(* IEC 61131-3 sources: Aqueous_Solutions/docs-authority/plc, 18 files *)

(* ---- PLC-CRYO.st ---- *)
(* AQS-CTL-004 X-CTL-04: control program source, generated by flow_graph/control/plc_programs.py *)
(* Basis: AQS-CTL-001 INSTRUMENT_INDEX.csv, AQS-CTL-002 control architecture, graph set-points. *)
(* PLC-CRYO: CPU redundant pair; IO counts AI 36 AO 1 DI 19 DO 6 (modules per AQS-CTL-002, 16-channel, 20 % spare) *)
PROGRAM PLC_CRYO_CTRL
VAR
  (* 100 ms cyclic task per AQS-CTL-002 *)
  CRYO_AHU_COND_CONDENSABLEFT-01_PV : REAL ;  (* S70 normal 0.00 L/h )
  CRYO_AHU_COND_CONDENSABLEPT-01_PV : REAL ;  (* no design pressure on the graph )
  CRYO_AHU_COND_CONDENSABLETE-01_PV : REAL ;  (* band by service )
  CRYO_AHUFT-01_PV : REAL ;  (* S56 normal 0.00 L/h )
  CRYO_AHUFT-02_PV : REAL ;  (* S68 normal 4.27 L/h )
  CRYO_AHUFT-03_PV : REAL ;  (* S86 normal 0.00 L/h )
  CRYO_AHUFT-04_PV : REAL ;  (* IA-HVAC-COND normal 2.81 L/h )
  CRYO_AHUPT-01_PV : REAL ;  (* no design pressure on the graph )
  CRYO_AHUTE-01_PV : REAL ;  (* band by service )
  CRYO_ASUPT-01_PV : REAL ;  (* design 18.0 kPa g )
  CRYO_ASUTE-01_PV : REAL ;  (* band by service )
  CRYO_CO2PT-01_PV : REAL ;  (* design 2200.0 kPa g )
  CRYO_CO2TE-01_PV : REAL ;  (* design T 25 C )
  CRYO_DED_COOLPT-01_PV : REAL ;  (* no design pressure on the graph )
  CRYO_DED_COOLTE-01_PV : REAL ;  (* band by service )
  CRYO_H2PT-01_PV : REAL ;  (* design 22000.0 kPa g )
  CRYO_H2TE-01_PV : REAL ;  (* design T 25 C )
  CRYO_N2PT-01_PV : REAL ;  (* no design pressure on the graph )
  CRYO_N2TE-01_PV : REAL ;  (* band by service )
  CRYO_O2PT-01_PV : REAL ;  (* design 22000.0 kPa g )
  CRYO_O2TE-01_PV : REAL ;  (* design T 25 C )
  CRYO_HX_Q4PT-01_PV : REAL ;  (* no design pressure on the graph )
  CRYO_HX_Q4TE-01_PV : REAL ;  (* band by service )
  H2O_ELYZFT-01_PV : REAL ;  (* IA-ELY-H2 normal 0.43 L/h )
  H2O_ELYZFT-02_PV : REAL ;  (* IA-ELY-O2 normal 3.42 L/h )
  H2O_ELYZLT-01_PV : REAL ;  (* A-M-182 liquid height )
  H2O_ELYZPT-01_PV : REAL ;  (* design 990.0 kPa g )
  H2O_ELYZTE-01_PV : REAL ;  (* band by service )
  PROD_MEOHLT-01_PV : REAL ;  (* A-M-182 liquid height )
  PROD_MEOHPT-01_PV : REAL ;  (* no design pressure on the graph )
  PROD_MEOHTE-01_PV : REAL ;  (* band by service )
  PROD_O2PT-01_PV : REAL ;  (* no design pressure on the graph )
  PROD_O2TE-01_PV : REAL ;  (* band by service )
  AIR_RECEIVERPT-01_PV : REAL ;  (* no design pressure on the graph )
  AIR_RECEIVERTE-01_PV : REAL ;  (* band by service )
  PROD_MEOHFT-01_PV : REAL ;  (* methanol product: IA-MEOH-PROD 28.15 kg/d (1.50 L/h at 792 kg/m3) )
END_VAR

  (* FLOW control loop - set-point from the graph basis *)
  CRYO_AHU_COND_CONDENSABLEFT-01_SP := 0.0 ;  (* graph basis: S70 normal 0.00 L/h )
  FB_PI_CRYO_AHU_COND_CONDENSABLEFT-01( PV := CRYO_AHU_COND_CONDENSABLEFT-01_PV, SP := CRYO_AHU_COND_CONDENSABLEFT-01_SP );  (* PI per AQS-CTL-002; GAIN/KI entered at commissioning from the step test (AQS-COM-001 sec. 3), anti-windup clamp per this FB *)
  CRYO_AHU_COND_CONDENSABLEFT-01_ALARM_HI := 0.0 ;  (* expected-zero state: any positive PV alarms )

  (* PRESSURE monitoring block - indication, no set-point invented )
  FB_AI_CRYO_AHU_COND_CONDENSABLEPT-01( PV := CRYO_AHU_COND_CONDENSABLEPT-01_PV );
  CRYO_AHU_COND_CONDENSABLEPT-01_ALARM_HI := 9.0 ;  (* 90 % of span, registered LSH convention )

  (* TEMPERATURE monitoring block - indication, no set-point invented )
  FB_AI_CRYO_AHU_COND_CONDENSABLETE-01( PV := CRYO_AHU_COND_CONDENSABLETE-01_PV );
  CRYO_AHU_COND_CONDENSABLETE-01_ALARM_HI := 45.0 ;  (* 90 % of span, registered LSH convention )

  (* FLOW control loop - set-point from the graph basis *)
  CRYO_AHUFT-01_SP := 0.0 ;  (* graph basis: S56 normal 0.00 L/h )
  FB_PI_CRYO_AHUFT-01( PV := CRYO_AHUFT-01_PV, SP := CRYO_AHUFT-01_SP );  (* PI per AQS-CTL-002; GAIN/KI entered at commissioning from the step test (AQS-COM-001 sec. 3), anti-windup clamp per this FB *)
  CRYO_AHUFT-01_ALARM_HI := 0.0 ;  (* expected-zero state: any positive PV alarms )

  (* FLOW control loop - set-point from the graph basis *)
  CRYO_AHUFT-02_SP := 4.27 ;  (* graph basis: S68 normal 4.27 L/h )
  FB_PI_CRYO_AHUFT-02( PV := CRYO_AHUFT-02_PV, SP := CRYO_AHUFT-02_SP );  (* PI per AQS-CTL-002; GAIN/KI entered at commissioning from the step test (AQS-COM-001 sec. 3), anti-windup clamp per this FB *)
  CRYO_AHUFT-02_ALARM_HI := 4.697 ;  (* SP x 1.1 margin, A-M-188 margin class *)
  CRYO_AHUFT-02_ALARM_LO := 3.8429999999999995 ;

  (* FLOW control loop - set-point from the graph basis *)
  CRYO_AHUFT-03_SP := 0.0 ;  (* graph basis: S86 normal 0.00 L/h )
  FB_PI_CRYO_AHUFT-03( PV := CRYO_AHUFT-03_PV, SP := CRYO_AHUFT-03_SP );  (* PI per AQS-CTL-002; GAIN/KI entered at commissioning from the step test (AQS-COM-001 sec. 3), anti-windup clamp per this FB *)
  CRYO_AHUFT-03_ALARM_HI := 0.0 ;  (* expected-zero state: any positive PV alarms )

  (* FLOW control loop - set-point from the graph basis *)
  CRYO_AHUFT-04_SP := 2.81 ;  (* graph basis: IA-HVAC-COND normal 2.81 L/h )
  FB_PI_CRYO_AHUFT-04( PV := CRYO_AHUFT-04_PV, SP := CRYO_AHUFT-04_SP );  (* PI per AQS-CTL-002; GAIN/KI entered at commissioning from the step test (AQS-COM-001 sec. 3), anti-windup clamp per this FB *)
  CRYO_AHUFT-04_ALARM_HI := 3.091 ;  (* SP x 1.1 margin, A-M-188 margin class *)
  CRYO_AHUFT-04_ALARM_LO := 2.529 ;

  (* PRESSURE monitoring block - indication, no set-point invented )
  FB_AI_CRYO_AHUPT-01( PV := CRYO_AHUPT-01_PV );
  CRYO_AHUPT-01_ALARM_HI := 9.0 ;  (* 90 % of span, registered LSH convention )

  (* TEMPERATURE monitoring block - indication, no set-point invented )
  FB_AI_CRYO_AHUTE-01( PV := CRYO_AHUTE-01_PV );
  CRYO_AHUTE-01_ALARM_HI := 45.0 ;  (* 90 % of span, registered LSH convention )

  (* PRESSURE control loop - set-point from the graph basis *)
  CRYO_ASUPT-01_SP := 18.0 ;  (* graph basis: design 18.0 kPa g )
  FB_PI_CRYO_ASUPT-01( PV := CRYO_ASUPT-01_PV, SP := CRYO_ASUPT-01_SP );  (* PI per AQS-CTL-002; GAIN/KI entered at commissioning from the step test (AQS-COM-001 sec. 3), anti-windup clamp per this FB *)
  CRYO_ASUPT-01_ALARM_HI := 19.8 ;  (* SP x 1.1 margin, A-M-188 margin class *)
  CRYO_ASUPT-01_ALARM_LO := 16.2 ;

  (* TEMPERATURE monitoring block - indication, no set-point invented )
  FB_AI_CRYO_ASUTE-01( PV := CRYO_ASUTE-01_PV );
  CRYO_ASUTE-01_ALARM_HI := 45.0 ;  (* 90 % of span, registered LSH convention )

  (* PRESSURE control loop - set-point from the graph basis *)
  CRYO_CO2PT-01_SP := 2200.0 ;  (* graph basis: design 2200.0 kPa g )
  FB_PI_CRYO_CO2PT-01( PV := CRYO_CO2PT-01_PV, SP := CRYO_CO2PT-01_SP );  (* PI per AQS-CTL-002; GAIN/KI entered at commissioning from the step test (AQS-COM-001 sec. 3), anti-windup clamp per this FB *)
  CRYO_CO2PT-01_ALARM_HI := 2420.0 ;  (* SP x 1.1 margin, A-M-188 margin class *)
  CRYO_CO2PT-01_ALARM_LO := 1980.0 ;

  (* TEMPERATURE control loop - set-point from the graph basis *)
  CRYO_CO2TE-01_SP := 25.0 ;  (* graph basis: design T 25 C )
  FB_PI_CRYO_CO2TE-01( PV := CRYO_CO2TE-01_PV, SP := CRYO_CO2TE-01_SP );  (* PI per AQS-CTL-002; GAIN/KI entered at commissioning from the step test (AQS-COM-001 sec. 3), anti-windup clamp per this FB *)
  CRYO_CO2TE-01_ALARM_HI := 27.500000000000004 ;  (* SP x 1.1 margin, A-M-188 margin class *)
  CRYO_CO2TE-01_ALARM_LO := 22.5 ;

  (* PRESSURE monitoring block - indication, no set-point invented )
  FB_AI_CRYO_DED_COOLPT-01( PV := CRYO_DED_COOLPT-01_PV );
  CRYO_DED_COOLPT-01_ALARM_HI := 9.0 ;  (* 90 % of span, registered LSH convention )

  (* TEMPERATURE monitoring block - indication, no set-point invented )
  FB_AI_CRYO_DED_COOLTE-01( PV := CRYO_DED_COOLTE-01_PV );
  CRYO_DED_COOLTE-01_ALARM_HI := 45.0 ;  (* 90 % of span, registered LSH convention )

  (* PRESSURE control loop - set-point from the graph basis *)
  CRYO_H2PT-01_SP := 22000.0 ;  (* graph basis: design 22000.0 kPa g )
  FB_PI_CRYO_H2PT-01( PV := CRYO_H2PT-01_PV, SP := CRYO_H2PT-01_SP );  (* PI per AQS-CTL-002; GAIN/KI entered at commissioning from the step test (AQS-COM-001 sec. 3), anti-windup clamp per this FB *)
  CRYO_H2PT-01_ALARM_HI := 24200.000000000004 ;  (* SP x 1.1 margin, A-M-188 margin class *)
  CRYO_H2PT-01_ALARM_LO := 19800.0 ;

  (* TEMPERATURE control loop - set-point from the graph basis *)
  CRYO_H2TE-01_SP := 25.0 ;  (* graph basis: design T 25 C )
  FB_PI_CRYO_H2TE-01( PV := CRYO_H2TE-01_PV, SP := CRYO_H2TE-01_SP );  (* PI per AQS-CTL-002; GAIN/KI entered at commissioning from the step test (AQS-COM-001 sec. 3), anti-windup clamp per this FB *)
  CRYO_H2TE-01_ALARM_HI := 27.500000000000004 ;  (* SP x 1.1 margin, A-M-188 margin class *)
  CRYO_H2TE-01_ALARM_LO := 22.5 ;

  (* PRESSURE monitoring block - indication, no set-point invented )
  FB_AI_CRYO_N2PT-01( PV := CRYO_N2PT-01_PV );
  CRYO_N2PT-01_ALARM_HI := 9.0 ;  (* 90 % of span, registered LSH convention )

  (* TEMPERATURE monitoring block - indication, no set-point invented )
  FB_AI_CRYO_N2TE-01( PV := CRYO_N2TE-01_PV );
  CRYO_N2TE-01_ALARM_HI := 45.0 ;  (* 90 % of span, registered LSH convention )

  (* PRESSURE control loop - set-point from the graph basis *)
  CRYO_O2PT-01_SP := 22000.0 ;  (* graph basis: design 22000.0 kPa g )
  FB_PI_CRYO_O2PT-01( PV := CRYO_O2PT-01_PV, SP := CRYO_O2PT-01_SP );  (* PI per AQS-CTL-002; GAIN/KI entered at commissioning from the step test (AQS-COM-001 sec. 3), anti-windup clamp per this FB *)
  CRYO_O2PT-01_ALARM_HI := 24200.000000000004 ;  (* SP x 1.1 margin, A-M-188 margin class *)
  CRYO_O2PT-01_ALARM_LO := 19800.0 ;

  (* TEMPERATURE control loop - set-point from the graph basis *)
  CRYO_O2TE-01_SP := 25.0 ;  (* graph basis: design T 25 C )
  FB_PI_CRYO_O2TE-01( PV := CRYO_O2TE-01_PV, SP := CRYO_O2TE-01_SP );  (* PI per AQS-CTL-002; GAIN/KI entered at commissioning from the step test (AQS-COM-001 sec. 3), anti-windup clamp per this FB *)
  CRYO_O2TE-01_ALARM_HI := 27.500000000000004 ;  (* SP x 1.1 margin, A-M-188 margin class *)
  CRYO_O2TE-01_ALARM_LO := 22.5 ;

  (* PRESSURE monitoring block - indication, no set-point invented )
  FB_AI_CRYO_HX_Q4PT-01( PV := CRYO_HX_Q4PT-01_PV );
  CRYO_HX_Q4PT-01_ALARM_HI := 9.0 ;  (* 90 % of span, registered LSH convention )

  (* TEMPERATURE monitoring block - indication, no set-point invented )
  FB_AI_CRYO_HX_Q4TE-01( PV := CRYO_HX_Q4TE-01_PV );
  CRYO_HX_Q4TE-01_ALARM_HI := 45.0 ;  (* 90 % of span, registered LSH convention )

  (* FLOW control loop - set-point from the graph basis *)
  H2O_ELYZFT-01_SP := 0.43 ;  (* graph basis: IA-ELY-H2 normal 0.43 L/h )
  FB_PI_H2O_ELYZFT-01( PV := H2O_ELYZFT-01_PV, SP := H2O_ELYZFT-01_SP );  (* PI per AQS-CTL-002; GAIN/KI entered at commissioning from the step test (AQS-COM-001 sec. 3), anti-windup clamp per this FB *)
  H2O_ELYZFT-01_ALARM_HI := 0.47300000000000003 ;  (* SP x 1.1 margin, A-M-188 margin class *)
  H2O_ELYZFT-01_ALARM_LO := 0.387 ;

  (* FLOW control loop - set-point from the graph basis *)
  H2O_ELYZFT-02_SP := 3.42 ;  (* graph basis: IA-ELY-O2 normal 3.42 L/h )
  FB_PI_H2O_ELYZFT-02( PV := H2O_ELYZFT-02_PV, SP := H2O_ELYZFT-02_SP );  (* PI per AQS-CTL-002; GAIN/KI entered at commissioning from the step test (AQS-COM-001 sec. 3), anti-windup clamp per this FB *)
  H2O_ELYZFT-02_ALARM_HI := 3.762 ;  (* SP x 1.1 margin, A-M-188 margin class *)
  H2O_ELYZFT-02_ALARM_LO := 3.078 ;

  (* LEVEL monitoring block - indication, no set-point invented )
  FB_AI_H2O_ELYZLT-01( PV := H2O_ELYZLT-01_PV );
  H2O_ELYZLT-01_ALARM_HI := 90.0 ;  (* 90 % of span, registered LSH convention )

  (* PRESSURE control loop - set-point from the graph basis *)
  H2O_ELYZPT-01_SP := 990.0 ;  (* graph basis: design 990.0 kPa g )
  FB_PI_H2O_ELYZPT-01( PV := H2O_ELYZPT-01_PV, SP := H2O_ELYZPT-01_SP );  (* PI per AQS-CTL-002; GAIN/KI entered at commissioning from the step test (AQS-COM-001 sec. 3), anti-windup clamp per this FB *)
  H2O_ELYZPT-01_ALARM_HI := 1089.0 ;  (* SP x 1.1 margin, A-M-188 margin class *)
  H2O_ELYZPT-01_ALARM_LO := 891.0 ;

  (* TEMPERATURE monitoring block - indication, no set-point invented )
  FB_AI_H2O_ELYZTE-01( PV := H2O_ELYZTE-01_PV );
  H2O_ELYZTE-01_ALARM_HI := 135.0 ;  (* 90 % of span, registered LSH convention )

  (* LEVEL monitoring block - indication, no set-point invented )
  FB_AI_PROD_MEOHLT-01( PV := PROD_MEOHLT-01_PV );
  PROD_MEOHLT-01_ALARM_HI := 90.0 ;  (* 90 % of span, registered LSH convention )

  (* PRESSURE monitoring block - indication, no set-point invented )
  FB_AI_PROD_MEOHPT-01( PV := PROD_MEOHPT-01_PV );
  PROD_MEOHPT-01_ALARM_HI := 9.0 ;  (* 90 % of span, registered LSH convention )

  (* TEMPERATURE monitoring block - indication, no set-point invented )
  FB_AI_PROD_MEOHTE-01( PV := PROD_MEOHTE-01_PV );
  PROD_MEOHTE-01_ALARM_HI := 135.0 ;  (* 90 % of span, registered LSH convention )

  (* PRESSURE monitoring block - indication, no set-point invented )
  FB_AI_PROD_O2PT-01( PV := PROD_O2PT-01_PV );
  PROD_O2PT-01_ALARM_HI := 9.0 ;  (* 90 % of span, registered LSH convention )

  (* TEMPERATURE monitoring block - indication, no set-point invented )
  FB_AI_PROD_O2TE-01( PV := PROD_O2TE-01_PV );
  PROD_O2TE-01_ALARM_HI := 135.0 ;  (* 90 % of span, registered LSH convention )

  (* PRESSURE monitoring block - indication, no set-point invented )
  FB_AI_AIR_RECEIVERPT-01( PV := AIR_RECEIVERPT-01_PV );
  AIR_RECEIVERPT-01_ALARM_HI := 9.0 ;  (* 90 % of span, registered LSH convention )

  (* TEMPERATURE monitoring block - indication, no set-point invented )
  FB_AI_AIR_RECEIVERTE-01( PV := AIR_RECEIVERTE-01_PV );
  AIR_RECEIVERTE-01_ALARM_HI := 135.0 ;  (* 90 % of span, registered LSH convention )

  (* FLOW monitoring block - indication, no set-point invented )
  FB_AI_PROD_MEOHFT-01( PV := PROD_MEOHFT-01_PV );
  PROD_MEOHFT-01_ALARM_HI := 4.5 ;  (* 90 % of span, registered LSH convention )

END_PROGRAM

(* ---- PLC-DIGESTER.st ---- *)
(* AQS-CTL-004 X-CTL-04: control program source, generated by flow_graph/control/plc_programs.py *)
(* Basis: AQS-CTL-001 INSTRUMENT_INDEX.csv, AQS-CTL-002 control architecture, graph set-points. *)
(* PLC-DIGESTER: CPU single; IO counts AI 135 AO 3 DI 121 DO 25 (modules per AQS-CTL-002, 16-channel, 20 % spare) *)
PROGRAM PLC_DIGESTER_CTRL
VAR
  (* 100 ms cyclic task per AQS-CTL-002 *)
  S13_CLASS_TREATPT-01_PV : REAL ;  (* no design pressure on the graph )
  S13_CLASS_TREATTE-01_PV : REAL ;  (* band by service )
  BMED_ACIDFT-01_PV : REAL ;  (* IA-BMED-01 normal 0.05 L/h )
  BMED_ACIDFT-02_PV : REAL ;  (* S09 normal 0.39 L/h )
  BMED_ACIDFT-03_PV : REAL ;  (* IA-EVAP_ACID-FEED normal 54.37 L/h )
  BMED_ACIDLT-01_PV : REAL ;  (* A-M-182 liquid height )
  BMED_ACIDPT-01_PV : REAL ;  (* no design pressure on the graph )
  BMED_ACIDTE-01_PV : REAL ;  (* band by service )
  BMED_BASEFT-01_PV : REAL ;  (* IA-BMED-02 normal 0.01 L/h )
  BMED_BASEFT-02_PV : REAL ;  (* IA-EVAP_BASE-FEED normal 54.24 L/h )
  BMED_BASEFT-03_PV : REAL ;  (* IA-VS-NAOH normal 0.00 L/h )
  BMED_BASELT-01_PV : REAL ;  (* A-M-182 liquid height )
  BMED_BASEPT-01_PV : REAL ;  (* no design pressure on the graph )
  BMED_BASETE-01_PV : REAL ;  (* band by service )
  CRUFT-01_PV : REAL ;  (* CRU_TO_VDF normal 0.01 L/h )
  CRUFT-02_PV : REAL ;  (* CRU_TO_TFE normal 0.01 L/h )
  CRUFT-03_PV : REAL ;  (* IA-CRU-01 normal 1.15 L/h )
  CRULT-01_PV : REAL ;  (* A-M-182 liquid height )
  CRUPT-01_PV : REAL ;  (* no design pressure on the graph )
  CRUTE-01_PV : REAL ;  (* band by service )
  EVAP_ACIDFT-01_PV : REAL ;  (* IA-ACID-01 normal 18.32 L/h )
  EVAP_ACIDFT-02_PV : REAL ;  (* IA-EVAP_ACID-COND normal 36.05 L/h )
  EVAP_ACIDFT-03_PV : REAL ;  (* IA-EVAP_ACID-VENT normal 0.00 L/h )
  EVAP_ACIDLT-01_PV : REAL ;  (* A-M-182 liquid height )
  EVAP_ACIDPT-01_PV : REAL ;  (* design 100.0 kPa g )
  EVAP_ACIDTE-01_PV : REAL ;  (* band by service )
  EVAP_ACID_VSFT-01_PV : REAL ;  (* IA-VS-SPENT normal 0.00 L/h )
  EVAP_ACID_VSFT-02_PV : REAL ;  (* IA-VS-OFF normal 0.00 L/h )
  EVAP_ACID_VSLT-01_PV : REAL ;  (* A-M-182 liquid height )
  EVAP_ACID_VSPT-01_PV : REAL ;  (* no design pressure on the graph )
  EVAP_ACID_VSTE-01_PV : REAL ;  (* band by service )
  EVAP_BASEFT-01_PV : REAL ;  (* IA-BASE-01 normal 0.92 L/h )
  EVAP_BASEFT-02_PV : REAL ;  (* IA-BASE-PPT normal 20.10 L/h )
  EVAP_BASEFT-03_PV : REAL ;  (* IA-EVAP_BASE-COND normal 33.80 L/h )
  EVAP_BASELT-01_PV : REAL ;  (* A-M-182 liquid height )
  EVAP_BASEPT-01_PV : REAL ;  (* design 100.0 kPa g )
  EVAP_BASETE-01_PV : REAL ;  (* band by service )
  FLOAT_SINKFT-01_PV : REAL ;  (* IA-WET-FLOAT-01 normal 13.68 L/h )
  FLOAT_SINKFT-02_PV : REAL ;  (* IA-PLAST-01 normal 1.38 L/h )
  FLOAT_SINKLT-01_PV : REAL ;  (* A-M-182 liquid height )
  FLOAT_SINKPT-01_PV : REAL ;  (* no design pressure on the graph )
  FLOAT_SINKTE-01_PV : REAL ;  (* band by service )
  F_RECOVERFT-01_PV : REAL ;  (* F_RECOVER_TO_HF_GEN normal 0.06 L/h )
  F_RECOVERLT-01_PV : REAL ;  (* A-M-182 liquid height )
  F_RECOVERPT-01_PV : REAL ;  (* no design pressure on the graph )
  F_RECOVERTE-01_PV : REAL ;  (* band by service )
  LI_RECOVERLT-01_PV : REAL ;  (* A-M-182 liquid height )
  LI_RECOVERPT-01_PV : REAL ;  (* no design pressure on the graph )
  LI_RECOVERTE-01_PV : REAL ;  (* band by service )
  POLISH_BANKFT-01_PV : REAL ;  (* IA-POL-01 normal 0.00 L/h )
  POLISH_BANKFT-02_PV : REAL ;  (* IA-POL-02 normal 164.40 L/h )
  POLISH_BANKFT-03_PV : REAL ;  (* POLISH_TO_LI normal 0.02 L/h )
  POLISH_BANKLT-01_PV : REAL ;  (* A-M-182 liquid height )
  POLISH_BANKPT-01_PV : REAL ;  (* no design pressure on the graph )
  POLISH_BANKTE-01_PV : REAL ;  (* band by service )
  P_CALT-01_PV : REAL ;  (* A-M-182 liquid height )
  P_CAPT-01_PV : REAL ;  (* no design pressure on the graph )
  P_CATE-01_PV : REAL ;  (* band by service )
  SALT_FEEDPT-01_PV : REAL ;  (* no design pressure on the graph )
  SALT_FEEDTE-01_PV : REAL ;  (* band by service )
  EW_1FT-01_PV : REAL ;  (* IA-EW-01 normal 178.66 L/h )
  EW_1FT-02_PV : REAL ;  (* IA-HDR-H2-01 normal 0.00 L/h )
  EW_1FT-03_PV : REAL ;  (* IA-HX8 normal 0.19 L/h )
  EW_1FT-04_PV : REAL ;  (* IA-EW1-H2 normal 0.00 L/h )
  EW_1FT-05_PV : REAL ;  (* IA-EW1-CL2 normal 0.00 L/h )
  EW_1LT-01_PV : REAL ;  (* A-M-182 liquid height )
  EW_1PT-01_PV : REAL ;  (* no design pressure on the graph )
  EW_1TE-01_PV : REAL ;  (* band by service )
  EW_2FT-01_PV : REAL ;  (* IA-EW-02 normal 178.66 L/h )
  EW_2FT-02_PV : REAL ;  (* IA-HDR-H2-03 normal 0.00 L/h )
  EW_2FT-03_PV : REAL ;  (* IA-EW2-H2 normal 0.00 L/h )
  EW_2FT-04_PV : REAL ;  (* IA-EW2-CL2 normal 0.00 L/h )
  EW_2LT-01_PV : REAL ;  (* A-M-182 liquid height )
  EW_2PT-01_PV : REAL ;  (* no design pressure on the graph )
  EW_2TE-01_PV : REAL ;  (* band by service )
  EW_9FT-01_PV : REAL ;  (* IA-EW-09 normal 173.46 L/h )
  EW_9FT-02_PV : REAL ;  (* IA-HDR-H2-04 normal 0.00 L/h )
  EW_9FT-03_PV : REAL ;  (* EW9_LIQUOR_TO_MO normal 0.00 L/h )
  EW_9FT-04_PV : REAL ;  (* IA-EW9-CL2 normal 0.25 L/h )
  EW_9LT-01_PV : REAL ;  (* A-M-182 liquid height )
  EW_9PT-01_PV : REAL ;  (* no design pressure on the graph )
  EW_9TE-01_PV : REAL ;  (* band by service )
  LEACH_CSTR_1LT-01_PV : REAL ;  (* A-M-182 liquid height )
  LEACH_CSTR_1PT-01_PV : REAL ;  (* no design pressure on the graph )
  LEACH_CSTR_1TE-01_PV : REAL ;  (* band by service )
  EW_3FT-01_PV : REAL ;  (* IA-EW-03 normal 177.64 L/h )
  EW_3FT-02_PV : REAL ;  (* IA-EW3-CL2 normal 1.01 L/h )
  EW_3FT-03_PV : REAL ;  (* IA-EW3-H2B normal 0.00 L/h )
  EW_3LT-01_PV : REAL ;  (* A-M-182 liquid height )
  EW_3PT-01_PV : REAL ;  (* no design pressure on the graph )
  EW_3TE-01_PV : REAL ;  (* band by service )
  EW_4FT-01_PV : REAL ;  (* IA-EW-10 normal 177.55 L/h )
  EW_4FT-02_PV : REAL ;  (* IA-EW4-H2 normal 0.00 L/h )
  EW_4FT-03_PV : REAL ;  (* IA-EW4-N2 normal 0.02 L/h )
  EW_4FT-04_PV : REAL ;  (* IA-EW4-CL2 normal 0.08 L/h )
  EW_4LT-01_PV : REAL ;  (* A-M-182 liquid height )
  EW_4PT-01_PV : REAL ;  (* no design pressure on the graph )
  EW_4TE-01_PV : REAL ;  (* band by service )
  EW_5FT-01_PV : REAL ;  (* IA-EW-05 normal 177.41 L/h )
  EW_5FT-02_PV : REAL ;  (* IA-EW5-CL2 normal 0.14 L/h )
  EW_5FT-03_PV : REAL ;  (* IA-EW5-H2B normal 0.00 L/h )
  EW_5LT-01_PV : REAL ;  (* A-M-182 liquid height )
  EW_5PT-01_PV : REAL ;  (* no design pressure on the graph )
  EW_5TE-01_PV : REAL ;  (* band by service )
  EW_6FT-01_PV : REAL ;  (* IA-EW-06 normal 177.14 L/h )
  EW_6FT-02_PV : REAL ;  (* IA-EW6-CL2 normal 0.27 L/h )
  EW_6FT-03_PV : REAL ;  (* IA-EW6-H2B normal 0.00 L/h )
  EW_6LT-01_PV : REAL ;  (* A-M-182 liquid height )
  EW_6PT-01_PV : REAL ;  (* no design pressure on the graph )
  EW_6TE-01_PV : REAL ;  (* band by service )
  EW_7FT-01_PV : REAL ;  (* IA-EW-07 normal 174.26 L/h )
  EW_7FT-02_PV : REAL ;  (* IA-EW7-CL2 normal 1.80 L/h )
  EW_7FT-03_PV : REAL ;  (* IA-EW7-H2B normal 0.01 L/h )
  EW_7LT-01_PV : REAL ;  (* A-M-182 liquid height )
  EW_7PT-01_PV : REAL ;  (* no design pressure on the graph )
  EW_7TE-01_PV : REAL ;  (* band by service )
  EW_8FT-01_PV : REAL ;  (* IA-EW-08 normal 174.12 L/h )
  EW_8FT-02_PV : REAL ;  (* IA-EW8-CL2 normal 0.14 L/h )
  EW_8FT-03_PV : REAL ;  (* IA-EW8-H2B normal 0.00 L/h )
  EW_8LT-01_PV : REAL ;  (* A-M-182 liquid height )
  EW_8PT-01_PV : REAL ;  (* no design pressure on the graph )
  EW_8TE-01_PV : REAL ;  (* band by service )
  HX8PT-01_PV : REAL ;  (* no design pressure on the graph )
  HX8TE-01_PV : REAL ;  (* band by service )
  NAOH_PLANTLT-01_PV : REAL ;  (* A-M-182 liquid height )
  NAOH_PLANTPT-01_PV : REAL ;  (* no design pressure on the graph )
  NAOH_PLANTTE-01_PV : REAL ;  (* band by service )
  CONTINUOUS_RECYCLELT-01_PV : REAL ;  (* A-M-182 liquid height )
  CONTINUOUS_RECYCLEPT-01_PV : REAL ;  (* no design pressure on the graph )
  CONTINUOUS_RECYCLETE-01_PV : REAL ;  (* band by service )
  EVAP_ACID_VSAE-01_PV : REAL ;  (* scrub liquor: NaOH 2 M bleed IA-VS-NAOH 0.5 g/d )
  EVAP_ACID_VSAE-02_PV : REAL ;  (* acid-gas breakthrough watch: IA-VS-OFF 0.029 kg/d scrubbed vent )
  EVAP_ACIDTE-90 : BOOL ;  (* SIF watch input, routed to the safety CPU pair (AQS-CTL-003) *)
  EVAP_ACID_VSTE-90 : BOOL ;  (* SIF watch input, routed to the safety CPU pair (AQS-CTL-003) *)
  EVAP_BASETE-90 : BOOL ;  (* SIF watch input, routed to the safety CPU pair (AQS-CTL-003) *)
END_VAR

  (* PRESSURE monitoring block - indication, no set-point invented )
  FB_AI_S13_CLASS_TREATPT-01( PV := S13_CLASS_TREATPT-01_PV );
  S13_CLASS_TREATPT-01_ALARM_HI := 9.0 ;  (* 90 % of span, registered LSH convention )

  (* TEMPERATURE monitoring block - indication, no set-point invented )
  FB_AI_S13_CLASS_TREATTE-01( PV := S13_CLASS_TREATTE-01_PV );
  S13_CLASS_TREATTE-01_ALARM_HI := 135.0 ;  (* 90 % of span, registered LSH convention )

  (* FLOW control loop - set-point from the graph basis *)
  BMED_ACIDFT-01_SP := 0.05 ;  (* graph basis: IA-BMED-01 normal 0.05 L/h )
  FB_PI_BMED_ACIDFT-01( PV := BMED_ACIDFT-01_PV, SP := BMED_ACIDFT-01_SP );  (* PI per AQS-CTL-002; GAIN/KI entered at commissioning from the step test (AQS-COM-001 sec. 3), anti-windup clamp per this FB *)
  BMED_ACIDFT-01_ALARM_HI := 0.05500000000000001 ;  (* SP x 1.1 margin, A-M-188 margin class *)
  BMED_ACIDFT-01_ALARM_LO := 0.045000000000000005 ;

  (* FLOW control loop - set-point from the graph basis *)
  BMED_ACIDFT-02_SP := 0.39 ;  (* graph basis: S09 normal 0.39 L/h )
  FB_PI_BMED_ACIDFT-02( PV := BMED_ACIDFT-02_PV, SP := BMED_ACIDFT-02_SP );  (* PI per AQS-CTL-002; GAIN/KI entered at commissioning from the step test (AQS-COM-001 sec. 3), anti-windup clamp per this FB *)
  BMED_ACIDFT-02_ALARM_HI := 0.42900000000000005 ;  (* SP x 1.1 margin, A-M-188 margin class *)
  BMED_ACIDFT-02_ALARM_LO := 0.35100000000000003 ;

  (* FLOW control loop - set-point from the graph basis *)
  BMED_ACIDFT-03_SP := 54.37 ;  (* graph basis: IA-EVAP_ACID-FEED normal 54.37 L/h )
  FB_PI_BMED_ACIDFT-03( PV := BMED_ACIDFT-03_PV, SP := BMED_ACIDFT-03_SP );  (* PI per AQS-CTL-002; GAIN/KI entered at commissioning from the step test (AQS-COM-001 sec. 3), anti-windup clamp per this FB *)
  BMED_ACIDFT-03_ALARM_HI := 59.807 ;  (* SP x 1.1 margin, A-M-188 margin class *)
  BMED_ACIDFT-03_ALARM_LO := 48.933 ;

  (* LEVEL monitoring block - indication, no set-point invented )
  FB_AI_BMED_ACIDLT-01( PV := BMED_ACIDLT-01_PV );
  BMED_ACIDLT-01_ALARM_HI := 90.0 ;  (* 90 % of span, registered LSH convention )

  (* PRESSURE monitoring block - indication, no set-point invented )
  FB_AI_BMED_ACIDPT-01( PV := BMED_ACIDPT-01_PV );
  BMED_ACIDPT-01_ALARM_HI := 9.0 ;  (* 90 % of span, registered LSH convention )

  (* TEMPERATURE monitoring block - indication, no set-point invented )
  FB_AI_BMED_ACIDTE-01( PV := BMED_ACIDTE-01_PV );
  BMED_ACIDTE-01_ALARM_HI := 135.0 ;  (* 90 % of span, registered LSH convention )

  (* FLOW control loop - set-point from the graph basis *)
  BMED_BASEFT-01_SP := 0.01 ;  (* graph basis: IA-BMED-02 normal 0.01 L/h )
  FB_PI_BMED_BASEFT-01( PV := BMED_BASEFT-01_PV, SP := BMED_BASEFT-01_SP );  (* PI per AQS-CTL-002; GAIN/KI entered at commissioning from the step test (AQS-COM-001 sec. 3), anti-windup clamp per this FB *)
  BMED_BASEFT-01_ALARM_HI := 0.011000000000000001 ;  (* SP x 1.1 margin, A-M-188 margin class *)
  BMED_BASEFT-01_ALARM_LO := 0.009000000000000001 ;

  (* FLOW control loop - set-point from the graph basis *)
  BMED_BASEFT-02_SP := 54.24 ;  (* graph basis: IA-EVAP_BASE-FEED normal 54.24 L/h )
  FB_PI_BMED_BASEFT-02( PV := BMED_BASEFT-02_PV, SP := BMED_BASEFT-02_SP );  (* PI per AQS-CTL-002; GAIN/KI entered at commissioning from the step test (AQS-COM-001 sec. 3), anti-windup clamp per this FB *)
  BMED_BASEFT-02_ALARM_HI := 59.66400000000001 ;  (* SP x 1.1 margin, A-M-188 margin class *)
  BMED_BASEFT-02_ALARM_LO := 48.816 ;

  (* FLOW control loop - set-point from the graph basis *)
  BMED_BASEFT-03_SP := 0.0 ;  (* graph basis: IA-VS-NAOH normal 0.00 L/h )
  FB_PI_BMED_BASEFT-03( PV := BMED_BASEFT-03_PV, SP := BMED_BASEFT-03_SP );  (* PI per AQS-CTL-002; GAIN/KI entered at commissioning from the step test (AQS-COM-001 sec. 3), anti-windup clamp per this FB *)
  BMED_BASEFT-03_ALARM_HI := 0.0 ;  (* expected-zero state: any positive PV alarms )

  (* LEVEL monitoring block - indication, no set-point invented )
  FB_AI_BMED_BASELT-01( PV := BMED_BASELT-01_PV );
  BMED_BASELT-01_ALARM_HI := 90.0 ;  (* 90 % of span, registered LSH convention )

  (* PRESSURE monitoring block - indication, no set-point invented )
  FB_AI_BMED_BASEPT-01( PV := BMED_BASEPT-01_PV );
  BMED_BASEPT-01_ALARM_HI := 9.0 ;  (* 90 % of span, registered LSH convention )

  (* TEMPERATURE monitoring block - indication, no set-point invented )
  FB_AI_BMED_BASETE-01( PV := BMED_BASETE-01_PV );
  BMED_BASETE-01_ALARM_HI := 135.0 ;  (* 90 % of span, registered LSH convention )

  (* FLOW control loop - set-point from the graph basis *)
  CRUFT-01_SP := 0.01 ;  (* graph basis: CRU_TO_VDF normal 0.01 L/h )
  FB_PI_CRUFT-01( PV := CRUFT-01_PV, SP := CRUFT-01_SP );  (* PI per AQS-CTL-002; GAIN/KI entered at commissioning from the step test (AQS-COM-001 sec. 3), anti-windup clamp per this FB *)
  CRUFT-01_ALARM_HI := 0.011000000000000001 ;  (* SP x 1.1 margin, A-M-188 margin class *)
  CRUFT-01_ALARM_LO := 0.009000000000000001 ;

  (* FLOW control loop - set-point from the graph basis *)
  CRUFT-02_SP := 0.01 ;  (* graph basis: CRU_TO_TFE normal 0.01 L/h )
  FB_PI_CRUFT-02( PV := CRUFT-02_PV, SP := CRUFT-02_SP );  (* PI per AQS-CTL-002; GAIN/KI entered at commissioning from the step test (AQS-COM-001 sec. 3), anti-windup clamp per this FB *)
  CRUFT-02_ALARM_HI := 0.011000000000000001 ;  (* SP x 1.1 margin, A-M-188 margin class *)
  CRUFT-02_ALARM_LO := 0.009000000000000001 ;

  (* FLOW control loop - set-point from the graph basis *)
  CRUFT-03_SP := 1.15 ;  (* graph basis: IA-CRU-01 normal 1.15 L/h )
  FB_PI_CRUFT-03( PV := CRUFT-03_PV, SP := CRUFT-03_SP );  (* PI per AQS-CTL-002; GAIN/KI entered at commissioning from the step test (AQS-COM-001 sec. 3), anti-windup clamp per this FB *)
  CRUFT-03_ALARM_HI := 1.265 ;  (* SP x 1.1 margin, A-M-188 margin class *)
  CRUFT-03_ALARM_LO := 1.035 ;

  (* LEVEL monitoring block - indication, no set-point invented )
  FB_AI_CRULT-01( PV := CRULT-01_PV );
  CRULT-01_ALARM_HI := 90.0 ;  (* 90 % of span, registered LSH convention )

  (* PRESSURE monitoring block - indication, no set-point invented )
  FB_AI_CRUPT-01( PV := CRUPT-01_PV );
  CRUPT-01_ALARM_HI := 9.0 ;  (* 90 % of span, registered LSH convention )

  (* TEMPERATURE monitoring block - indication, no set-point invented )
  FB_AI_CRUTE-01( PV := CRUTE-01_PV );
  CRUTE-01_ALARM_HI := 135.0 ;  (* 90 % of span, registered LSH convention )

  (* FLOW control loop - set-point from the graph basis *)
  EVAP_ACIDFT-01_SP := 18.32 ;  (* graph basis: IA-ACID-01 normal 18.32 L/h )
  FB_PI_EVAP_ACIDFT-01( PV := EVAP_ACIDFT-01_PV, SP := EVAP_ACIDFT-01_SP );  (* PI per AQS-CTL-002; GAIN/KI entered at commissioning from the step test (AQS-COM-001 sec. 3), anti-windup clamp per this FB *)
  EVAP_ACIDFT-01_ALARM_HI := 20.152 ;  (* SP x 1.1 margin, A-M-188 margin class *)
  EVAP_ACIDFT-01_ALARM_LO := 16.488 ;

  (* FLOW control loop - set-point from the graph basis *)
  EVAP_ACIDFT-02_SP := 36.05 ;  (* graph basis: IA-EVAP_ACID-COND normal 36.05 L/h )
  FB_PI_EVAP_ACIDFT-02( PV := EVAP_ACIDFT-02_PV, SP := EVAP_ACIDFT-02_SP );  (* PI per AQS-CTL-002; GAIN/KI entered at commissioning from the step test (AQS-COM-001 sec. 3), anti-windup clamp per this FB *)
  EVAP_ACIDFT-02_ALARM_HI := 39.655 ;  (* SP x 1.1 margin, A-M-188 margin class *)
  EVAP_ACIDFT-02_ALARM_LO := 32.445 ;

  (* FLOW control loop - set-point from the graph basis *)
  EVAP_ACIDFT-03_SP := 0.0 ;  (* graph basis: IA-EVAP_ACID-VENT normal 0.00 L/h )
  FB_PI_EVAP_ACIDFT-03( PV := EVAP_ACIDFT-03_PV, SP := EVAP_ACIDFT-03_SP );  (* PI per AQS-CTL-002; GAIN/KI entered at commissioning from the step test (AQS-COM-001 sec. 3), anti-windup clamp per this FB *)
  EVAP_ACIDFT-03_ALARM_HI := 0.0 ;  (* expected-zero state: any positive PV alarms )

  (* LEVEL monitoring block - indication, no set-point invented )
  FB_AI_EVAP_ACIDLT-01( PV := EVAP_ACIDLT-01_PV );
  EVAP_ACIDLT-01_ALARM_HI := 90.0 ;  (* 90 % of span, registered LSH convention )

  (* PRESSURE control loop - set-point from the graph basis *)
  EVAP_ACIDPT-01_SP := 100.0 ;  (* graph basis: design 100.0 kPa g )
  FB_PI_EVAP_ACIDPT-01( PV := EVAP_ACIDPT-01_PV, SP := EVAP_ACIDPT-01_SP );  (* PI per AQS-CTL-002; GAIN/KI entered at commissioning from the step test (AQS-COM-001 sec. 3), anti-windup clamp per this FB *)
  EVAP_ACIDPT-01_ALARM_HI := 110.00000000000001 ;  (* SP x 1.1 margin, A-M-188 margin class *)
  EVAP_ACIDPT-01_ALARM_LO := 90.0 ;

  (* TEMPERATURE monitoring block - indication, no set-point invented )
  FB_AI_EVAP_ACIDTE-01( PV := EVAP_ACIDTE-01_PV );
  EVAP_ACIDTE-01_ALARM_HI := 540.0 ;  (* 90 % of span, registered LSH convention )

  (* FLOW control loop - set-point from the graph basis *)
  EVAP_ACID_VSFT-01_SP := 0.0 ;  (* graph basis: IA-VS-SPENT normal 0.00 L/h )
  FB_PI_EVAP_ACID_VSFT-01( PV := EVAP_ACID_VSFT-01_PV, SP := EVAP_ACID_VSFT-01_SP );  (* PI per AQS-CTL-002; GAIN/KI entered at commissioning from the step test (AQS-COM-001 sec. 3), anti-windup clamp per this FB *)
  EVAP_ACID_VSFT-01_ALARM_HI := 0.0 ;  (* expected-zero state: any positive PV alarms )

  (* FLOW control loop - set-point from the graph basis *)
  EVAP_ACID_VSFT-02_SP := 0.0 ;  (* graph basis: IA-VS-OFF normal 0.00 L/h )
  FB_PI_EVAP_ACID_VSFT-02( PV := EVAP_ACID_VSFT-02_PV, SP := EVAP_ACID_VSFT-02_SP );  (* PI per AQS-CTL-002; GAIN/KI entered at commissioning from the step test (AQS-COM-001 sec. 3), anti-windup clamp per this FB *)
  EVAP_ACID_VSFT-02_ALARM_HI := 0.0 ;  (* expected-zero state: any positive PV alarms )

  (* LEVEL monitoring block - indication, no set-point invented )
  FB_AI_EVAP_ACID_VSLT-01( PV := EVAP_ACID_VSLT-01_PV );
  EVAP_ACID_VSLT-01_ALARM_HI := 90.0 ;  (* 90 % of span, registered LSH convention )

  (* PRESSURE monitoring block - indication, no set-point invented )
  FB_AI_EVAP_ACID_VSPT-01( PV := EVAP_ACID_VSPT-01_PV );
  EVAP_ACID_VSPT-01_ALARM_HI := 9.0 ;  (* 90 % of span, registered LSH convention )

  (* TEMPERATURE monitoring block - indication, no set-point invented )
  FB_AI_EVAP_ACID_VSTE-01( PV := EVAP_ACID_VSTE-01_PV );
  EVAP_ACID_VSTE-01_ALARM_HI := 540.0 ;  (* 90 % of span, registered LSH convention )

  (* FLOW control loop - set-point from the graph basis *)
  EVAP_BASEFT-01_SP := 0.92 ;  (* graph basis: IA-BASE-01 normal 0.92 L/h )
  FB_PI_EVAP_BASEFT-01( PV := EVAP_BASEFT-01_PV, SP := EVAP_BASEFT-01_SP );  (* PI per AQS-CTL-002; GAIN/KI entered at commissioning from the step test (AQS-COM-001 sec. 3), anti-windup clamp per this FB *)
  EVAP_BASEFT-01_ALARM_HI := 1.0120000000000002 ;  (* SP x 1.1 margin, A-M-188 margin class *)
  EVAP_BASEFT-01_ALARM_LO := 0.8280000000000001 ;

  (* FLOW control loop - set-point from the graph basis *)
  EVAP_BASEFT-02_SP := 20.1 ;  (* graph basis: IA-BASE-PPT normal 20.10 L/h )
  FB_PI_EVAP_BASEFT-02( PV := EVAP_BASEFT-02_PV, SP := EVAP_BASEFT-02_SP );  (* PI per AQS-CTL-002; GAIN/KI entered at commissioning from the step test (AQS-COM-001 sec. 3), anti-windup clamp per this FB *)
  EVAP_BASEFT-02_ALARM_HI := 22.110000000000003 ;  (* SP x 1.1 margin, A-M-188 margin class *)
  EVAP_BASEFT-02_ALARM_LO := 18.090000000000003 ;

  (* FLOW control loop - set-point from the graph basis *)
  EVAP_BASEFT-03_SP := 33.8 ;  (* graph basis: IA-EVAP_BASE-COND normal 33.80 L/h )
  FB_PI_EVAP_BASEFT-03( PV := EVAP_BASEFT-03_PV, SP := EVAP_BASEFT-03_SP );  (* PI per AQS-CTL-002; GAIN/KI entered at commissioning from the step test (AQS-COM-001 sec. 3), anti-windup clamp per this FB *)
  EVAP_BASEFT-03_ALARM_HI := 37.18 ;  (* SP x 1.1 margin, A-M-188 margin class *)
  EVAP_BASEFT-03_ALARM_LO := 30.419999999999998 ;

  (* LEVEL monitoring block - indication, no set-point invented )
  FB_AI_EVAP_BASELT-01( PV := EVAP_BASELT-01_PV );
  EVAP_BASELT-01_ALARM_HI := 90.0 ;  (* 90 % of span, registered LSH convention )

  (* PRESSURE control loop - set-point from the graph basis *)
  EVAP_BASEPT-01_SP := 100.0 ;  (* graph basis: design 100.0 kPa g )
  FB_PI_EVAP_BASEPT-01( PV := EVAP_BASEPT-01_PV, SP := EVAP_BASEPT-01_SP );  (* PI per AQS-CTL-002; GAIN/KI entered at commissioning from the step test (AQS-COM-001 sec. 3), anti-windup clamp per this FB *)
  EVAP_BASEPT-01_ALARM_HI := 110.00000000000001 ;  (* SP x 1.1 margin, A-M-188 margin class *)
  EVAP_BASEPT-01_ALARM_LO := 90.0 ;

  (* TEMPERATURE monitoring block - indication, no set-point invented )
  FB_AI_EVAP_BASETE-01( PV := EVAP_BASETE-01_PV );
  EVAP_BASETE-01_ALARM_HI := 540.0 ;  (* 90 % of span, registered LSH convention )

  (* FLOW control loop - set-point from the graph basis *)
  FLOAT_SINKFT-01_SP := 13.68 ;  (* graph basis: IA-WET-FLOAT-01 normal 13.68 L/h )
  FB_PI_FLOAT_SINKFT-01( PV := FLOAT_SINKFT-01_PV, SP := FLOAT_SINKFT-01_SP );  (* PI per AQS-CTL-002; GAIN/KI entered at commissioning from the step test (AQS-COM-001 sec. 3), anti-windup clamp per this FB *)
  FLOAT_SINKFT-01_ALARM_HI := 15.048 ;  (* SP x 1.1 margin, A-M-188 margin class *)
  FLOAT_SINKFT-01_ALARM_LO := 12.312 ;

  (* FLOW control loop - set-point from the graph basis *)
  FLOAT_SINKFT-02_SP := 1.38 ;  (* graph basis: IA-PLAST-01 normal 1.38 L/h )
  FB_PI_FLOAT_SINKFT-02( PV := FLOAT_SINKFT-02_PV, SP := FLOAT_SINKFT-02_SP );  (* PI per AQS-CTL-002; GAIN/KI entered at commissioning from the step test (AQS-COM-001 sec. 3), anti-windup clamp per this FB *)
  FLOAT_SINKFT-02_ALARM_HI := 1.518 ;  (* SP x 1.1 margin, A-M-188 margin class *)
  FLOAT_SINKFT-02_ALARM_LO := 1.242 ;

  (* LEVEL monitoring block - indication, no set-point invented )
  FB_AI_FLOAT_SINKLT-01( PV := FLOAT_SINKLT-01_PV );
  FLOAT_SINKLT-01_ALARM_HI := 90.0 ;  (* 90 % of span, registered LSH convention )

  (* PRESSURE monitoring block - indication, no set-point invented )
  FB_AI_FLOAT_SINKPT-01( PV := FLOAT_SINKPT-01_PV );
  FLOAT_SINKPT-01_ALARM_HI := 9.0 ;  (* 90 % of span, registered LSH convention )

  (* TEMPERATURE monitoring block - indication, no set-point invented )
  FB_AI_FLOAT_SINKTE-01( PV := FLOAT_SINKTE-01_PV );
  FLOAT_SINKTE-01_ALARM_HI := 135.0 ;  (* 90 % of span, registered LSH convention )

  (* FLOW control loop - set-point from the graph basis *)
  F_RECOVERFT-01_SP := 0.06 ;  (* graph basis: F_RECOVER_TO_HF_GEN normal 0.06 L/h )
  FB_PI_F_RECOVERFT-01( PV := F_RECOVERFT-01_PV, SP := F_RECOVERFT-01_SP );  (* PI per AQS-CTL-002; GAIN/KI entered at commissioning from the step test (AQS-COM-001 sec. 3), anti-windup clamp per this FB *)
  F_RECOVERFT-01_ALARM_HI := 0.066 ;  (* SP x 1.1 margin, A-M-188 margin class *)
  F_RECOVERFT-01_ALARM_LO := 0.054 ;

  (* LEVEL monitoring block - indication, no set-point invented )
  FB_AI_F_RECOVERLT-01( PV := F_RECOVERLT-01_PV );
  F_RECOVERLT-01_ALARM_HI := 90.0 ;  (* 90 % of span, registered LSH convention )

  (* PRESSURE monitoring block - indication, no set-point invented )
  FB_AI_F_RECOVERPT-01( PV := F_RECOVERPT-01_PV );
  F_RECOVERPT-01_ALARM_HI := 9.0 ;  (* 90 % of span, registered LSH convention )

  (* TEMPERATURE monitoring block - indication, no set-point invented )
  FB_AI_F_RECOVERTE-01( PV := F_RECOVERTE-01_PV );
  F_RECOVERTE-01_ALARM_HI := 135.0 ;  (* 90 % of span, registered LSH convention )

  (* LEVEL monitoring block - indication, no set-point invented )
  FB_AI_LI_RECOVERLT-01( PV := LI_RECOVERLT-01_PV );
  LI_RECOVERLT-01_ALARM_HI := 90.0 ;  (* 90 % of span, registered LSH convention )

  (* PRESSURE monitoring block - indication, no set-point invented )
  FB_AI_LI_RECOVERPT-01( PV := LI_RECOVERPT-01_PV );
  LI_RECOVERPT-01_ALARM_HI := 9.0 ;  (* 90 % of span, registered LSH convention )

  (* TEMPERATURE monitoring block - indication, no set-point invented )
  FB_AI_LI_RECOVERTE-01( PV := LI_RECOVERTE-01_PV );
  LI_RECOVERTE-01_ALARM_HI := 135.0 ;  (* 90 % of span, registered LSH convention )

  (* FLOW control loop - set-point from the graph basis *)
  POLISH_BANKFT-01_SP := 0.0 ;  (* graph basis: IA-POL-01 normal 0.00 L/h )
  FB_PI_POLISH_BANKFT-01( PV := POLISH_BANKFT-01_PV, SP := POLISH_BANKFT-01_SP );  (* PI per AQS-CTL-002; GAIN/KI entered at commissioning from the step test (AQS-COM-001 sec. 3), anti-windup clamp per this FB *)
  POLISH_BANKFT-01_ALARM_HI := 0.0 ;  (* expected-zero state: any positive PV alarms )

  (* FLOW control loop - set-point from the graph basis *)
  POLISH_BANKFT-02_SP := 164.4 ;  (* graph basis: IA-POL-02 normal 164.40 L/h )
  FB_PI_POLISH_BANKFT-02( PV := POLISH_BANKFT-02_PV, SP := POLISH_BANKFT-02_SP );  (* PI per AQS-CTL-002; GAIN/KI entered at commissioning from the step test (AQS-COM-001 sec. 3), anti-windup clamp per this FB *)
  POLISH_BANKFT-02_ALARM_HI := 180.84000000000003 ;  (* SP x 1.1 margin, A-M-188 margin class *)
  POLISH_BANKFT-02_ALARM_LO := 147.96 ;

  (* FLOW control loop - set-point from the graph basis *)
  POLISH_BANKFT-03_SP := 0.02 ;  (* graph basis: POLISH_TO_LI normal 0.02 L/h )
  FB_PI_POLISH_BANKFT-03( PV := POLISH_BANKFT-03_PV, SP := POLISH_BANKFT-03_SP );  (* PI per AQS-CTL-002; GAIN/KI entered at commissioning from the step test (AQS-COM-001 sec. 3), anti-windup clamp per this FB *)
  POLISH_BANKFT-03_ALARM_HI := 0.022000000000000002 ;  (* SP x 1.1 margin, A-M-188 margin class *)
  POLISH_BANKFT-03_ALARM_LO := 0.018000000000000002 ;

  (* LEVEL monitoring block - indication, no set-point invented )
  FB_AI_POLISH_BANKLT-01( PV := POLISH_BANKLT-01_PV );
  POLISH_BANKLT-01_ALARM_HI := 90.0 ;  (* 90 % of span, registered LSH convention )

  (* PRESSURE monitoring block - indication, no set-point invented )
  FB_AI_POLISH_BANKPT-01( PV := POLISH_BANKPT-01_PV );
  POLISH_BANKPT-01_ALARM_HI := 9.0 ;  (* 90 % of span, registered LSH convention )

  (* TEMPERATURE monitoring block - indication, no set-point invented )
  FB_AI_POLISH_BANKTE-01( PV := POLISH_BANKTE-01_PV );
  POLISH_BANKTE-01_ALARM_HI := 135.0 ;  (* 90 % of span, registered LSH convention )

  (* LEVEL monitoring block - indication, no set-point invented )
  FB_AI_P_CALT-01( PV := P_CALT-01_PV );
  P_CALT-01_ALARM_HI := 90.0 ;  (* 90 % of span, registered LSH convention )

  (* PRESSURE monitoring block - indication, no set-point invented )
  FB_AI_P_CAPT-01( PV := P_CAPT-01_PV );
  P_CAPT-01_ALARM_HI := 9.0 ;  (* 90 % of span, registered LSH convention )

  (* TEMPERATURE monitoring block - indication, no set-point invented )
  FB_AI_P_CATE-01( PV := P_CATE-01_PV );
  P_CATE-01_ALARM_HI := 135.0 ;  (* 90 % of span, registered LSH convention )

  (* PRESSURE monitoring block - indication, no set-point invented )
  FB_AI_SALT_FEEDPT-01( PV := SALT_FEEDPT-01_PV );
  SALT_FEEDPT-01_ALARM_HI := 9.0 ;  (* 90 % of span, registered LSH convention )

  (* TEMPERATURE monitoring block - indication, no set-point invented )
  FB_AI_SALT_FEEDTE-01( PV := SALT_FEEDTE-01_PV );
  SALT_FEEDTE-01_ALARM_HI := 135.0 ;  (* 90 % of span, registered LSH convention )

  (* FLOW control loop - set-point from the graph basis *)
  EW_1FT-01_SP := 178.66 ;  (* graph basis: IA-EW-01 normal 178.66 L/h )
  FB_PI_EW_1FT-01( PV := EW_1FT-01_PV, SP := EW_1FT-01_SP );  (* PI per AQS-CTL-002; GAIN/KI entered at commissioning from the step test (AQS-COM-001 sec. 3), anti-windup clamp per this FB *)
  EW_1FT-01_ALARM_HI := 196.526 ;  (* SP x 1.1 margin, A-M-188 margin class *)
  EW_1FT-01_ALARM_LO := 160.794 ;

  (* FLOW control loop - set-point from the graph basis *)
  EW_1FT-02_SP := 0.0 ;  (* graph basis: IA-HDR-H2-01 normal 0.00 L/h )
  FB_PI_EW_1FT-02( PV := EW_1FT-02_PV, SP := EW_1FT-02_SP );  (* PI per AQS-CTL-002; GAIN/KI entered at commissioning from the step test (AQS-COM-001 sec. 3), anti-windup clamp per this FB *)
  EW_1FT-02_ALARM_HI := 0.0 ;  (* expected-zero state: any positive PV alarms )

  (* FLOW control loop - set-point from the graph basis *)
  EW_1FT-03_SP := 0.19 ;  (* graph basis: IA-HX8 normal 0.19 L/h )
  FB_PI_EW_1FT-03( PV := EW_1FT-03_PV, SP := EW_1FT-03_SP );  (* PI per AQS-CTL-002; GAIN/KI entered at commissioning from the step test (AQS-COM-001 sec. 3), anti-windup clamp per this FB *)
  EW_1FT-03_ALARM_HI := 0.20900000000000002 ;  (* SP x 1.1 margin, A-M-188 margin class *)
  EW_1FT-03_ALARM_LO := 0.171 ;

  (* FLOW control loop - set-point from the graph basis *)
  EW_1FT-04_SP := 0.0 ;  (* graph basis: IA-EW1-H2 normal 0.00 L/h )
  FB_PI_EW_1FT-04( PV := EW_1FT-04_PV, SP := EW_1FT-04_SP );  (* PI per AQS-CTL-002; GAIN/KI entered at commissioning from the step test (AQS-COM-001 sec. 3), anti-windup clamp per this FB *)
  EW_1FT-04_ALARM_HI := 0.0 ;  (* expected-zero state: any positive PV alarms )

  (* FLOW control loop - set-point from the graph basis *)
  EW_1FT-05_SP := 0.0 ;  (* graph basis: IA-EW1-CL2 normal 0.00 L/h )
  FB_PI_EW_1FT-05( PV := EW_1FT-05_PV, SP := EW_1FT-05_SP );  (* PI per AQS-CTL-002; GAIN/KI entered at commissioning from the step test (AQS-COM-001 sec. 3), anti-windup clamp per this FB *)
  EW_1FT-05_ALARM_HI := 0.0 ;  (* expected-zero state: any positive PV alarms )

  (* LEVEL monitoring block - indication, no set-point invented )
  FB_AI_EW_1LT-01( PV := EW_1LT-01_PV );
  EW_1LT-01_ALARM_HI := 90.0 ;  (* 90 % of span, registered LSH convention )

  (* PRESSURE monitoring block - indication, no set-point invented )
  FB_AI_EW_1PT-01( PV := EW_1PT-01_PV );
  EW_1PT-01_ALARM_HI := 9.0 ;  (* 90 % of span, registered LSH convention )

  (* TEMPERATURE monitoring block - indication, no set-point invented )
  FB_AI_EW_1TE-01( PV := EW_1TE-01_PV );
  EW_1TE-01_ALARM_HI := 135.0 ;  (* 90 % of span, registered LSH convention )

  (* FLOW control loop - set-point from the graph basis *)
  EW_2FT-01_SP := 178.66 ;  (* graph basis: IA-EW-02 normal 178.66 L/h )
  FB_PI_EW_2FT-01( PV := EW_2FT-01_PV, SP := EW_2FT-01_SP );  (* PI per AQS-CTL-002; GAIN/KI entered at commissioning from the step test (AQS-COM-001 sec. 3), anti-windup clamp per this FB *)
  EW_2FT-01_ALARM_HI := 196.526 ;  (* SP x 1.1 margin, A-M-188 margin class *)
  EW_2FT-01_ALARM_LO := 160.794 ;

  (* FLOW control loop - set-point from the graph basis *)
  EW_2FT-02_SP := 0.0 ;  (* graph basis: IA-HDR-H2-03 normal 0.00 L/h )
  FB_PI_EW_2FT-02( PV := EW_2FT-02_PV, SP := EW_2FT-02_SP );  (* PI per AQS-CTL-002; GAIN/KI entered at commissioning from the step test (AQS-COM-001 sec. 3), anti-windup clamp per this FB *)
  EW_2FT-02_ALARM_HI := 0.0 ;  (* expected-zero state: any positive PV alarms )

  (* FLOW control loop - set-point from the graph basis *)
  EW_2FT-03_SP := 0.0 ;  (* graph basis: IA-EW2-H2 normal 0.00 L/h )
  FB_PI_EW_2FT-03( PV := EW_2FT-03_PV, SP := EW_2FT-03_SP );  (* PI per AQS-CTL-002; GAIN/KI entered at commissioning from the step test (AQS-COM-001 sec. 3), anti-windup clamp per this FB *)
  EW_2FT-03_ALARM_HI := 0.0 ;  (* expected-zero state: any positive PV alarms )

  (* FLOW control loop - set-point from the graph basis *)
  EW_2FT-04_SP := 0.0 ;  (* graph basis: IA-EW2-CL2 normal 0.00 L/h )
  FB_PI_EW_2FT-04( PV := EW_2FT-04_PV, SP := EW_2FT-04_SP );  (* PI per AQS-CTL-002; GAIN/KI entered at commissioning from the step test (AQS-COM-001 sec. 3), anti-windup clamp per this FB *)
  EW_2FT-04_ALARM_HI := 0.0 ;  (* expected-zero state: any positive PV alarms )

  (* LEVEL monitoring block - indication, no set-point invented )
  FB_AI_EW_2LT-01( PV := EW_2LT-01_PV );
  EW_2LT-01_ALARM_HI := 90.0 ;  (* 90 % of span, registered LSH convention )

  (* PRESSURE monitoring block - indication, no set-point invented )
  FB_AI_EW_2PT-01( PV := EW_2PT-01_PV );
  EW_2PT-01_ALARM_HI := 9.0 ;  (* 90 % of span, registered LSH convention )

  (* TEMPERATURE monitoring block - indication, no set-point invented )
  FB_AI_EW_2TE-01( PV := EW_2TE-01_PV );
  EW_2TE-01_ALARM_HI := 135.0 ;  (* 90 % of span, registered LSH convention )

  (* FLOW control loop - set-point from the graph basis *)
  EW_9FT-01_SP := 173.46 ;  (* graph basis: IA-EW-09 normal 173.46 L/h )
  FB_PI_EW_9FT-01( PV := EW_9FT-01_PV, SP := EW_9FT-01_SP );  (* PI per AQS-CTL-002; GAIN/KI entered at commissioning from the step test (AQS-COM-001 sec. 3), anti-windup clamp per this FB *)
  EW_9FT-01_ALARM_HI := 190.806 ;  (* SP x 1.1 margin, A-M-188 margin class *)
  EW_9FT-01_ALARM_LO := 156.114 ;

  (* FLOW control loop - set-point from the graph basis *)
  EW_9FT-02_SP := 0.0 ;  (* graph basis: IA-HDR-H2-04 normal 0.00 L/h )
  FB_PI_EW_9FT-02( PV := EW_9FT-02_PV, SP := EW_9FT-02_SP );  (* PI per AQS-CTL-002; GAIN/KI entered at commissioning from the step test (AQS-COM-001 sec. 3), anti-windup clamp per this FB *)
  EW_9FT-02_ALARM_HI := 0.0 ;  (* expected-zero state: any positive PV alarms )

  (* FLOW control loop - set-point from the graph basis *)
  EW_9FT-03_SP := 0.0 ;  (* graph basis: EW9_LIQUOR_TO_MO normal 0.00 L/h )
  FB_PI_EW_9FT-03( PV := EW_9FT-03_PV, SP := EW_9FT-03_SP );  (* PI per AQS-CTL-002; GAIN/KI entered at commissioning from the step test (AQS-COM-001 sec. 3), anti-windup clamp per this FB *)
  EW_9FT-03_ALARM_HI := 0.0 ;  (* expected-zero state: any positive PV alarms )

  (* FLOW control loop - set-point from the graph basis *)
  EW_9FT-04_SP := 0.25 ;  (* graph basis: IA-EW9-CL2 normal 0.25 L/h )
  FB_PI_EW_9FT-04( PV := EW_9FT-04_PV, SP := EW_9FT-04_SP );  (* PI per AQS-CTL-002; GAIN/KI entered at commissioning from the step test (AQS-COM-001 sec. 3), anti-windup clamp per this FB *)
  EW_9FT-04_ALARM_HI := 0.275 ;  (* SP x 1.1 margin, A-M-188 margin class *)
  EW_9FT-04_ALARM_LO := 0.225 ;

  (* LEVEL monitoring block - indication, no set-point invented )
  FB_AI_EW_9LT-01( PV := EW_9LT-01_PV );
  EW_9LT-01_ALARM_HI := 90.0 ;  (* 90 % of span, registered LSH convention )

  (* PRESSURE monitoring block - indication, no set-point invented )
  FB_AI_EW_9PT-01( PV := EW_9PT-01_PV );
  EW_9PT-01_ALARM_HI := 9.0 ;  (* 90 % of span, registered LSH convention )

  (* TEMPERATURE monitoring block - indication, no set-point invented )
  FB_AI_EW_9TE-01( PV := EW_9TE-01_PV );
  EW_9TE-01_ALARM_HI := 135.0 ;  (* 90 % of span, registered LSH convention )

  (* LEVEL monitoring block - indication, no set-point invented )
  FB_AI_LEACH_CSTR_1LT-01( PV := LEACH_CSTR_1LT-01_PV );
  LEACH_CSTR_1LT-01_ALARM_HI := 90.0 ;  (* 90 % of span, registered LSH convention )

  (* PRESSURE monitoring block - indication, no set-point invented )
  FB_AI_LEACH_CSTR_1PT-01( PV := LEACH_CSTR_1PT-01_PV );
  LEACH_CSTR_1PT-01_ALARM_HI := 9.0 ;  (* 90 % of span, registered LSH convention )

  (* TEMPERATURE monitoring block - indication, no set-point invented )
  FB_AI_LEACH_CSTR_1TE-01( PV := LEACH_CSTR_1TE-01_PV );
  LEACH_CSTR_1TE-01_ALARM_HI := 135.0 ;  (* 90 % of span, registered LSH convention )

  (* FLOW control loop - set-point from the graph basis *)
  EW_3FT-01_SP := 177.64 ;  (* graph basis: IA-EW-03 normal 177.64 L/h )
  FB_PI_EW_3FT-01( PV := EW_3FT-01_PV, SP := EW_3FT-01_SP );  (* PI per AQS-CTL-002; GAIN/KI entered at commissioning from the step test (AQS-COM-001 sec. 3), anti-windup clamp per this FB *)
  EW_3FT-01_ALARM_HI := 195.404 ;  (* SP x 1.1 margin, A-M-188 margin class *)
  EW_3FT-01_ALARM_LO := 159.876 ;

  (* FLOW control loop - set-point from the graph basis *)
  EW_3FT-02_SP := 1.01 ;  (* graph basis: IA-EW3-CL2 normal 1.01 L/h )
  FB_PI_EW_3FT-02( PV := EW_3FT-02_PV, SP := EW_3FT-02_SP );  (* PI per AQS-CTL-002; GAIN/KI entered at commissioning from the step test (AQS-COM-001 sec. 3), anti-windup clamp per this FB *)
  EW_3FT-02_ALARM_HI := 1.1110000000000002 ;  (* SP x 1.1 margin, A-M-188 margin class *)
  EW_3FT-02_ALARM_LO := 0.909 ;

  (* FLOW control loop - set-point from the graph basis *)
  EW_3FT-03_SP := 0.0 ;  (* graph basis: IA-EW3-H2B normal 0.00 L/h )
  FB_PI_EW_3FT-03( PV := EW_3FT-03_PV, SP := EW_3FT-03_SP );  (* PI per AQS-CTL-002; GAIN/KI entered at commissioning from the step test (AQS-COM-001 sec. 3), anti-windup clamp per this FB *)
  EW_3FT-03_ALARM_HI := 0.0 ;  (* expected-zero state: any positive PV alarms )

  (* LEVEL monitoring block - indication, no set-point invented )
  FB_AI_EW_3LT-01( PV := EW_3LT-01_PV );
  EW_3LT-01_ALARM_HI := 90.0 ;  (* 90 % of span, registered LSH convention )

  (* PRESSURE monitoring block - indication, no set-point invented )
  FB_AI_EW_3PT-01( PV := EW_3PT-01_PV );
  EW_3PT-01_ALARM_HI := 9.0 ;  (* 90 % of span, registered LSH convention )

  (* TEMPERATURE monitoring block - indication, no set-point invented )
  FB_AI_EW_3TE-01( PV := EW_3TE-01_PV );
  EW_3TE-01_ALARM_HI := 135.0 ;  (* 90 % of span, registered LSH convention )

  (* FLOW control loop - set-point from the graph basis *)
  EW_4FT-01_SP := 177.55 ;  (* graph basis: IA-EW-10 normal 177.55 L/h )
  FB_PI_EW_4FT-01( PV := EW_4FT-01_PV, SP := EW_4FT-01_SP );  (* PI per AQS-CTL-002; GAIN/KI entered at commissioning from the step test (AQS-COM-001 sec. 3), anti-windup clamp per this FB *)
  EW_4FT-01_ALARM_HI := 195.30500000000004 ;  (* SP x 1.1 margin, A-M-188 margin class *)
  EW_4FT-01_ALARM_LO := 159.79500000000002 ;

  (* FLOW control loop - set-point from the graph basis *)
  EW_4FT-02_SP := 0.0 ;  (* graph basis: IA-EW4-H2 normal 0.00 L/h )
  FB_PI_EW_4FT-02( PV := EW_4FT-02_PV, SP := EW_4FT-02_SP );  (* PI per AQS-CTL-002; GAIN/KI entered at commissioning from the step test (AQS-COM-001 sec. 3), anti-windup clamp per this FB *)
  EW_4FT-02_ALARM_HI := 0.0 ;  (* expected-zero state: any positive PV alarms )

  (* FLOW control loop - set-point from the graph basis *)
  EW_4FT-03_SP := 0.02 ;  (* graph basis: IA-EW4-N2 normal 0.02 L/h )
  FB_PI_EW_4FT-03( PV := EW_4FT-03_PV, SP := EW_4FT-03_SP );  (* PI per AQS-CTL-002; GAIN/KI entered at commissioning from the step test (AQS-COM-001 sec. 3), anti-windup clamp per this FB *)
  EW_4FT-03_ALARM_HI := 0.022000000000000002 ;  (* SP x 1.1 margin, A-M-188 margin class *)
  EW_4FT-03_ALARM_LO := 0.018000000000000002 ;

  (* FLOW control loop - set-point from the graph basis *)
  EW_4FT-04_SP := 0.08 ;  (* graph basis: IA-EW4-CL2 normal 0.08 L/h )
  FB_PI_EW_4FT-04( PV := EW_4FT-04_PV, SP := EW_4FT-04_SP );  (* PI per AQS-CTL-002; GAIN/KI entered at commissioning from the step test (AQS-COM-001 sec. 3), anti-windup clamp per this FB *)
  EW_4FT-04_ALARM_HI := 0.08800000000000001 ;  (* SP x 1.1 margin, A-M-188 margin class *)
  EW_4FT-04_ALARM_LO := 0.07200000000000001 ;

  (* LEVEL monitoring block - indication, no set-point invented )
  FB_AI_EW_4LT-01( PV := EW_4LT-01_PV );
  EW_4LT-01_ALARM_HI := 90.0 ;  (* 90 % of span, registered LSH convention )

  (* PRESSURE monitoring block - indication, no set-point invented )
  FB_AI_EW_4PT-01( PV := EW_4PT-01_PV );
  EW_4PT-01_ALARM_HI := 9.0 ;  (* 90 % of span, registered LSH convention )

  (* TEMPERATURE monitoring block - indication, no set-point invented )
  FB_AI_EW_4TE-01( PV := EW_4TE-01_PV );
  EW_4TE-01_ALARM_HI := 135.0 ;  (* 90 % of span, registered LSH convention )

  (* FLOW control loop - set-point from the graph basis *)
  EW_5FT-01_SP := 177.41 ;  (* graph basis: IA-EW-05 normal 177.41 L/h )
  FB_PI_EW_5FT-01( PV := EW_5FT-01_PV, SP := EW_5FT-01_SP );  (* PI per AQS-CTL-002; GAIN/KI entered at commissioning from the step test (AQS-COM-001 sec. 3), anti-windup clamp per this FB *)
  EW_5FT-01_ALARM_HI := 195.151 ;  (* SP x 1.1 margin, A-M-188 margin class *)
  EW_5FT-01_ALARM_LO := 159.669 ;

  (* FLOW control loop - set-point from the graph basis *)
  EW_5FT-02_SP := 0.14 ;  (* graph basis: IA-EW5-CL2 normal 0.14 L/h )
  FB_PI_EW_5FT-02( PV := EW_5FT-02_PV, SP := EW_5FT-02_SP );  (* PI per AQS-CTL-002; GAIN/KI entered at commissioning from the step test (AQS-COM-001 sec. 3), anti-windup clamp per this FB *)
  EW_5FT-02_ALARM_HI := 0.15400000000000003 ;  (* SP x 1.1 margin, A-M-188 margin class *)
  EW_5FT-02_ALARM_LO := 0.12600000000000003 ;

  (* FLOW control loop - set-point from the graph basis *)
  EW_5FT-03_SP := 0.0 ;  (* graph basis: IA-EW5-H2B normal 0.00 L/h )
  FB_PI_EW_5FT-03( PV := EW_5FT-03_PV, SP := EW_5FT-03_SP );  (* PI per AQS-CTL-002; GAIN/KI entered at commissioning from the step test (AQS-COM-001 sec. 3), anti-windup clamp per this FB *)
  EW_5FT-03_ALARM_HI := 0.0 ;  (* expected-zero state: any positive PV alarms )

  (* LEVEL monitoring block - indication, no set-point invented )
  FB_AI_EW_5LT-01( PV := EW_5LT-01_PV );
  EW_5LT-01_ALARM_HI := 90.0 ;  (* 90 % of span, registered LSH convention )

  (* PRESSURE monitoring block - indication, no set-point invented )
  FB_AI_EW_5PT-01( PV := EW_5PT-01_PV );
  EW_5PT-01_ALARM_HI := 9.0 ;  (* 90 % of span, registered LSH convention )

  (* TEMPERATURE monitoring block - indication, no set-point invented )
  FB_AI_EW_5TE-01( PV := EW_5TE-01_PV );
  EW_5TE-01_ALARM_HI := 135.0 ;  (* 90 % of span, registered LSH convention )

  (* FLOW control loop - set-point from the graph basis *)
  EW_6FT-01_SP := 177.14 ;  (* graph basis: IA-EW-06 normal 177.14 L/h )
  FB_PI_EW_6FT-01( PV := EW_6FT-01_PV, SP := EW_6FT-01_SP );  (* PI per AQS-CTL-002; GAIN/KI entered at commissioning from the step test (AQS-COM-001 sec. 3), anti-windup clamp per this FB *)
  EW_6FT-01_ALARM_HI := 194.854 ;  (* SP x 1.1 margin, A-M-188 margin class *)
  EW_6FT-01_ALARM_LO := 159.426 ;

  (* FLOW control loop - set-point from the graph basis *)
  EW_6FT-02_SP := 0.27 ;  (* graph basis: IA-EW6-CL2 normal 0.27 L/h )
  FB_PI_EW_6FT-02( PV := EW_6FT-02_PV, SP := EW_6FT-02_SP );  (* PI per AQS-CTL-002; GAIN/KI entered at commissioning from the step test (AQS-COM-001 sec. 3), anti-windup clamp per this FB *)
  EW_6FT-02_ALARM_HI := 0.29700000000000004 ;  (* SP x 1.1 margin, A-M-188 margin class *)
  EW_6FT-02_ALARM_LO := 0.24300000000000002 ;

  (* FLOW control loop - set-point from the graph basis *)
  EW_6FT-03_SP := 0.0 ;  (* graph basis: IA-EW6-H2B normal 0.00 L/h )
  FB_PI_EW_6FT-03( PV := EW_6FT-03_PV, SP := EW_6FT-03_SP );  (* PI per AQS-CTL-002; GAIN/KI entered at commissioning from the step test (AQS-COM-001 sec. 3), anti-windup clamp per this FB *)
  EW_6FT-03_ALARM_HI := 0.0 ;  (* expected-zero state: any positive PV alarms )

  (* LEVEL monitoring block - indication, no set-point invented )
  FB_AI_EW_6LT-01( PV := EW_6LT-01_PV );
  EW_6LT-01_ALARM_HI := 90.0 ;  (* 90 % of span, registered LSH convention )

  (* PRESSURE monitoring block - indication, no set-point invented )
  FB_AI_EW_6PT-01( PV := EW_6PT-01_PV );
  EW_6PT-01_ALARM_HI := 9.0 ;  (* 90 % of span, registered LSH convention )

  (* TEMPERATURE monitoring block - indication, no set-point invented )
  FB_AI_EW_6TE-01( PV := EW_6TE-01_PV );
  EW_6TE-01_ALARM_HI := 135.0 ;  (* 90 % of span, registered LSH convention )

  (* FLOW control loop - set-point from the graph basis *)
  EW_7FT-01_SP := 174.26 ;  (* graph basis: IA-EW-07 normal 174.26 L/h )
  FB_PI_EW_7FT-01( PV := EW_7FT-01_PV, SP := EW_7FT-01_SP );  (* PI per AQS-CTL-002; GAIN/KI entered at commissioning from the step test (AQS-COM-001 sec. 3), anti-windup clamp per this FB *)
  EW_7FT-01_ALARM_HI := 191.686 ;  (* SP x 1.1 margin, A-M-188 margin class *)
  EW_7FT-01_ALARM_LO := 156.834 ;

  (* FLOW control loop - set-point from the graph basis *)
  EW_7FT-02_SP := 1.8 ;  (* graph basis: IA-EW7-CL2 normal 1.80 L/h )
  FB_PI_EW_7FT-02( PV := EW_7FT-02_PV, SP := EW_7FT-02_SP );  (* PI per AQS-CTL-002; GAIN/KI entered at commissioning from the step test (AQS-COM-001 sec. 3), anti-windup clamp per this FB *)
  EW_7FT-02_ALARM_HI := 1.9800000000000002 ;  (* SP x 1.1 margin, A-M-188 margin class *)
  EW_7FT-02_ALARM_LO := 1.62 ;

  (* FLOW control loop - set-point from the graph basis *)
  EW_7FT-03_SP := 0.01 ;  (* graph basis: IA-EW7-H2B normal 0.01 L/h )
  FB_PI_EW_7FT-03( PV := EW_7FT-03_PV, SP := EW_7FT-03_SP );  (* PI per AQS-CTL-002; GAIN/KI entered at commissioning from the step test (AQS-COM-001 sec. 3), anti-windup clamp per this FB *)
  EW_7FT-03_ALARM_HI := 0.011000000000000001 ;  (* SP x 1.1 margin, A-M-188 margin class *)
  EW_7FT-03_ALARM_LO := 0.009000000000000001 ;

  (* LEVEL monitoring block - indication, no set-point invented )
  FB_AI_EW_7LT-01( PV := EW_7LT-01_PV );
  EW_7LT-01_ALARM_HI := 90.0 ;  (* 90 % of span, registered LSH convention )

  (* PRESSURE monitoring block - indication, no set-point invented )
  FB_AI_EW_7PT-01( PV := EW_7PT-01_PV );
  EW_7PT-01_ALARM_HI := 9.0 ;  (* 90 % of span, registered LSH convention )

  (* TEMPERATURE monitoring block - indication, no set-point invented )
  FB_AI_EW_7TE-01( PV := EW_7TE-01_PV );
  EW_7TE-01_ALARM_HI := 135.0 ;  (* 90 % of span, registered LSH convention )

  (* FLOW control loop - set-point from the graph basis *)
  EW_8FT-01_SP := 174.12 ;  (* graph basis: IA-EW-08 normal 174.12 L/h )
  FB_PI_EW_8FT-01( PV := EW_8FT-01_PV, SP := EW_8FT-01_SP );  (* PI per AQS-CTL-002; GAIN/KI entered at commissioning from the step test (AQS-COM-001 sec. 3), anti-windup clamp per this FB *)
  EW_8FT-01_ALARM_HI := 191.532 ;  (* SP x 1.1 margin, A-M-188 margin class *)
  EW_8FT-01_ALARM_LO := 156.708 ;

  (* FLOW control loop - set-point from the graph basis *)
  EW_8FT-02_SP := 0.14 ;  (* graph basis: IA-EW8-CL2 normal 0.14 L/h )
  FB_PI_EW_8FT-02( PV := EW_8FT-02_PV, SP := EW_8FT-02_SP );  (* PI per AQS-CTL-002; GAIN/KI entered at commissioning from the step test (AQS-COM-001 sec. 3), anti-windup clamp per this FB *)
  EW_8FT-02_ALARM_HI := 0.15400000000000003 ;  (* SP x 1.1 margin, A-M-188 margin class *)
  EW_8FT-02_ALARM_LO := 0.12600000000000003 ;

  (* FLOW control loop - set-point from the graph basis *)
  EW_8FT-03_SP := 0.0 ;  (* graph basis: IA-EW8-H2B normal 0.00 L/h )
  FB_PI_EW_8FT-03( PV := EW_8FT-03_PV, SP := EW_8FT-03_SP );  (* PI per AQS-CTL-002; GAIN/KI entered at commissioning from the step test (AQS-COM-001 sec. 3), anti-windup clamp per this FB *)
  EW_8FT-03_ALARM_HI := 0.0 ;  (* expected-zero state: any positive PV alarms )

  (* LEVEL monitoring block - indication, no set-point invented )
  FB_AI_EW_8LT-01( PV := EW_8LT-01_PV );
  EW_8LT-01_ALARM_HI := 90.0 ;  (* 90 % of span, registered LSH convention )

  (* PRESSURE monitoring block - indication, no set-point invented )
  FB_AI_EW_8PT-01( PV := EW_8PT-01_PV );
  EW_8PT-01_ALARM_HI := 9.0 ;  (* 90 % of span, registered LSH convention )

  (* TEMPERATURE monitoring block - indication, no set-point invented )
  FB_AI_EW_8TE-01( PV := EW_8TE-01_PV );
  EW_8TE-01_ALARM_HI := 135.0 ;  (* 90 % of span, registered LSH convention )

  (* PRESSURE monitoring block - indication, no set-point invented )
  FB_AI_HX8PT-01( PV := HX8PT-01_PV );
  HX8PT-01_ALARM_HI := 9.0 ;  (* 90 % of span, registered LSH convention )

  (* TEMPERATURE monitoring block - indication, no set-point invented )
  FB_AI_HX8TE-01( PV := HX8TE-01_PV );
  HX8TE-01_ALARM_HI := 135.0 ;  (* 90 % of span, registered LSH convention )

  (* LEVEL monitoring block - indication, no set-point invented )
  FB_AI_NAOH_PLANTLT-01( PV := NAOH_PLANTLT-01_PV );
  NAOH_PLANTLT-01_ALARM_HI := 90.0 ;  (* 90 % of span, registered LSH convention )

  (* PRESSURE monitoring block - indication, no set-point invented )
  FB_AI_NAOH_PLANTPT-01( PV := NAOH_PLANTPT-01_PV );
  NAOH_PLANTPT-01_ALARM_HI := 9.0 ;  (* 90 % of span, registered LSH convention )

  (* TEMPERATURE monitoring block - indication, no set-point invented )
  FB_AI_NAOH_PLANTTE-01( PV := NAOH_PLANTTE-01_PV );
  NAOH_PLANTTE-01_ALARM_HI := 135.0 ;  (* 90 % of span, registered LSH convention )

  (* LEVEL monitoring block - indication, no set-point invented )
  FB_AI_CONTINUOUS_RECYCLELT-01( PV := CONTINUOUS_RECYCLELT-01_PV );
  CONTINUOUS_RECYCLELT-01_ALARM_HI := 90.0 ;  (* 90 % of span, registered LSH convention )

  (* PRESSURE monitoring block - indication, no set-point invented )
  FB_AI_CONTINUOUS_RECYCLEPT-01( PV := CONTINUOUS_RECYCLEPT-01_PV );
  CONTINUOUS_RECYCLEPT-01_ALARM_HI := 9.0 ;  (* 90 % of span, registered LSH convention )

  (* TEMPERATURE monitoring block - indication, no set-point invented )
  FB_AI_CONTINUOUS_RECYCLETE-01( PV := CONTINUOUS_RECYCLETE-01_PV );
  CONTINUOUS_RECYCLETE-01_ALARM_HI := 135.0 ;  (* 90 % of span, registered LSH convention )

  (* PH monitoring block - indication, no set-point invented )
  FB_AI_EVAP_ACID_VSAE-01( PV := EVAP_ACID_VSAE-01_PV );
  EVAP_ACID_VSAE-01_ALARM_HI := 12.6 ;  (* 90 % of span, registered LSH convention )

  (* ORP monitoring block - indication, no set-point invented )
  FB_AI_EVAP_ACID_VSAE-02( PV := EVAP_ACID_VSAE-02_PV );
  EVAP_ACID_VSAE-02_ALARM_HI := 900.0 ;  (* 90 % of span, registered LSH convention )

  (* SIF watch passthrough, no action in the basic program )
  SIF_WATCH_EVAP_ACIDTE-90 := EVAP_ACIDTE-90 ;  (* to safety CPU pair, AQS-CTL-003 )

  (* SIF watch passthrough, no action in the basic program )
  SIF_WATCH_EVAP_ACID_VSTE-90 := EVAP_ACID_VSTE-90 ;  (* to safety CPU pair, AQS-CTL-003 )

  (* SIF watch passthrough, no action in the basic program )
  SIF_WATCH_EVAP_BASETE-90 := EVAP_BASETE-90 ;  (* to safety CPU pair, AQS-CTL-003 )

END_PROGRAM

(* ---- PLC-ELEC.st ---- *)
(* AQS-CTL-004 X-CTL-04: control program source, generated by flow_graph/control/plc_programs.py *)
(* Basis: AQS-CTL-001 INSTRUMENT_INDEX.csv, AQS-CTL-002 control architecture, graph set-points. *)
(* PLC-ELEC: CPU redundant pair; IO counts AI 29 AO 17 DI 445 DO 108 (modules per AQS-CTL-002, 16-channel, 20 % spare) *)
PROGRAM PLC_ELEC_CTRL
VAR
  (* 100 ms cyclic task per AQS-CTL-002 *)
  ZNBR2FT-01_PV : REAL ;  (* S69 normal 33.48 L/h )
  ZNBR2FT-02_PV : REAL ;  (* IA-ZNBR-BD normal 0.33 L/h )
  ZNBR2FT-03_PV : REAL ;  (* IA-ZNBR-HEAT normal 1.98 L/h )
  ZNBR2FT-04_PV : REAL ;  (* IA-ZNBR-H2 normal 0.03 L/h )
  ZNBR2LT-01_PV : REAL ;  (* A-M-182 liquid height )
  ZNBR2PT-01_PV : REAL ;  (* no design pressure on the graph )
  ZNBR2TE-01_PV : REAL ;  (* band by service )
  BACKUP_GENLT-01_PV : REAL ;  (* A-M-182 liquid height )
  BACKUP_GENPT-01_PV : REAL ;  (* no design pressure on the graph )
  BACKUP_GENTE-01_PV : REAL ;  (* band by service )
  SOL_ARK_60KPT-01_PV : REAL ;  (* no design pressure on the graph )
  SOL_ARK_60KTE-01_PV : REAL ;  (* band by service )
  LOAD_AGGPT-01_PV : REAL ;  (* no design pressure on the graph )
  LOAD_AGGTE-01_PV : REAL ;  (* band by service )
  FUEL_CELLFT-01_PV : REAL ;  (* S52 normal 1.79 L/h )
  FUEL_CELLFT-02_PV : REAL ;  (* IA-FC-FIX normal 0.00 L/h )
  FUEL_CELLFT-03_PV : REAL ;  (* IA-FC-LEACH normal 0.01 L/h )
  FUEL_CELLPT-01_PV : REAL ;  (* no design pressure on the graph )
  FUEL_CELLTE-01_PV : REAL ;  (* band by service )
  PV_ARRAYPT-01_PV : REAL ;  (* no design pressure on the graph )
  PV_ARRAYTE-01_PV : REAL ;  (* band by service )
  RECTIFIERPT-01_PV : REAL ;  (* no design pressure on the graph )
  RECTIFIERTE-01_PV : REAL ;  (* band by service )
  ZNBR2_BR2_REGENFT-01_PV : REAL ;  (* S69B normal 33.48 L/h )
  ZNBR2_BR2_REGENLT-01_PV : REAL ;  (* A-M-182 liquid height )
  ZNBR2_BR2_REGENPT-01_PV : REAL ;  (* no design pressure on the graph )
  ZNBR2_BR2_REGENTE-01_PV : REAL ;  (* band by service )
  EXT_HALLTE-01_PV : REAL ;  (* hall air: SF-EXT_HALL 68.28 kW electrical feed (ventilation watch) )
  LIO_BATPT-01_PV : REAL ;  (* pack enclosure pressure watch on the sealed storage (X-LOC-10 placeholder; A-M-4 )
END_VAR

  (* FLOW control loop - set-point from the graph basis *)
  ZNBR2FT-01_SP := 33.48 ;  (* graph basis: S69 normal 33.48 L/h )
  FB_PI_ZNBR2FT-01( PV := ZNBR2FT-01_PV, SP := ZNBR2FT-01_SP );  (* PI per AQS-CTL-002; GAIN/KI entered at commissioning from the step test (AQS-COM-001 sec. 3), anti-windup clamp per this FB *)
  ZNBR2FT-01_ALARM_HI := 36.828 ;  (* SP x 1.1 margin, A-M-188 margin class *)
  ZNBR2FT-01_ALARM_LO := 30.131999999999998 ;

  (* FLOW control loop - set-point from the graph basis *)
  ZNBR2FT-02_SP := 0.33 ;  (* graph basis: IA-ZNBR-BD normal 0.33 L/h )
  FB_PI_ZNBR2FT-02( PV := ZNBR2FT-02_PV, SP := ZNBR2FT-02_SP );  (* PI per AQS-CTL-002; GAIN/KI entered at commissioning from the step test (AQS-COM-001 sec. 3), anti-windup clamp per this FB *)
  ZNBR2FT-02_ALARM_HI := 0.36300000000000004 ;  (* SP x 1.1 margin, A-M-188 margin class *)
  ZNBR2FT-02_ALARM_LO := 0.29700000000000004 ;

  (* FLOW control loop - set-point from the graph basis *)
  ZNBR2FT-03_SP := 1.98 ;  (* graph basis: IA-ZNBR-HEAT normal 1.98 L/h )
  FB_PI_ZNBR2FT-03( PV := ZNBR2FT-03_PV, SP := ZNBR2FT-03_SP );  (* PI per AQS-CTL-002; GAIN/KI entered at commissioning from the step test (AQS-COM-001 sec. 3), anti-windup clamp per this FB *)
  ZNBR2FT-03_ALARM_HI := 2.178 ;  (* SP x 1.1 margin, A-M-188 margin class *)
  ZNBR2FT-03_ALARM_LO := 1.782 ;

  (* FLOW control loop - set-point from the graph basis *)
  ZNBR2FT-04_SP := 0.03 ;  (* graph basis: IA-ZNBR-H2 normal 0.03 L/h )
  FB_PI_ZNBR2FT-04( PV := ZNBR2FT-04_PV, SP := ZNBR2FT-04_SP );  (* PI per AQS-CTL-002; GAIN/KI entered at commissioning from the step test (AQS-COM-001 sec. 3), anti-windup clamp per this FB *)
  ZNBR2FT-04_ALARM_HI := 0.033 ;  (* SP x 1.1 margin, A-M-188 margin class *)
  ZNBR2FT-04_ALARM_LO := 0.027 ;

  (* LEVEL monitoring block - indication, no set-point invented )
  FB_AI_ZNBR2LT-01( PV := ZNBR2LT-01_PV );
  ZNBR2LT-01_ALARM_HI := 90.0 ;  (* 90 % of span, registered LSH convention )

  (* PRESSURE monitoring block - indication, no set-point invented )
  FB_AI_ZNBR2PT-01( PV := ZNBR2PT-01_PV );
  ZNBR2PT-01_ALARM_HI := 9.0 ;  (* 90 % of span, registered LSH convention )

  (* TEMPERATURE monitoring block - indication, no set-point invented )
  FB_AI_ZNBR2TE-01( PV := ZNBR2TE-01_PV );
  ZNBR2TE-01_ALARM_HI := 135.0 ;  (* 90 % of span, registered LSH convention )

  (* LEVEL monitoring block - indication, no set-point invented )
  FB_AI_BACKUP_GENLT-01( PV := BACKUP_GENLT-01_PV );
  BACKUP_GENLT-01_ALARM_HI := 90.0 ;  (* 90 % of span, registered LSH convention )

  (* PRESSURE monitoring block - indication, no set-point invented )
  FB_AI_BACKUP_GENPT-01( PV := BACKUP_GENPT-01_PV );
  BACKUP_GENPT-01_ALARM_HI := 9.0 ;  (* 90 % of span, registered LSH convention )

  (* TEMPERATURE monitoring block - indication, no set-point invented )
  FB_AI_BACKUP_GENTE-01( PV := BACKUP_GENTE-01_PV );
  BACKUP_GENTE-01_ALARM_HI := 135.0 ;  (* 90 % of span, registered LSH convention )

  (* PRESSURE monitoring block - indication, no set-point invented )
  FB_AI_SOL_ARK_60KPT-01( PV := SOL_ARK_60KPT-01_PV );
  SOL_ARK_60KPT-01_ALARM_HI := 9.0 ;  (* 90 % of span, registered LSH convention )

  (* TEMPERATURE monitoring block - indication, no set-point invented )
  FB_AI_SOL_ARK_60KTE-01( PV := SOL_ARK_60KTE-01_PV );
  SOL_ARK_60KTE-01_ALARM_HI := 135.0 ;  (* 90 % of span, registered LSH convention )

  (* PRESSURE monitoring block - indication, no set-point invented )
  FB_AI_LOAD_AGGPT-01( PV := LOAD_AGGPT-01_PV );
  LOAD_AGGPT-01_ALARM_HI := 9.0 ;  (* 90 % of span, registered LSH convention )

  (* TEMPERATURE monitoring block - indication, no set-point invented )
  FB_AI_LOAD_AGGTE-01( PV := LOAD_AGGTE-01_PV );
  LOAD_AGGTE-01_ALARM_HI := 135.0 ;  (* 90 % of span, registered LSH convention )

  (* FLOW control loop - set-point from the graph basis *)
  FUEL_CELLFT-01_SP := 1.79 ;  (* graph basis: S52 normal 1.79 L/h )
  FB_PI_FUEL_CELLFT-01( PV := FUEL_CELLFT-01_PV, SP := FUEL_CELLFT-01_SP );  (* PI per AQS-CTL-002; GAIN/KI entered at commissioning from the step test (AQS-COM-001 sec. 3), anti-windup clamp per this FB *)
  FUEL_CELLFT-01_ALARM_HI := 1.9690000000000003 ;  (* SP x 1.1 margin, A-M-188 margin class *)
  FUEL_CELLFT-01_ALARM_LO := 1.611 ;

  (* FLOW control loop - set-point from the graph basis *)
  FUEL_CELLFT-02_SP := 0.0 ;  (* graph basis: IA-FC-FIX normal 0.00 L/h )
  FB_PI_FUEL_CELLFT-02( PV := FUEL_CELLFT-02_PV, SP := FUEL_CELLFT-02_SP );  (* PI per AQS-CTL-002; GAIN/KI entered at commissioning from the step test (AQS-COM-001 sec. 3), anti-windup clamp per this FB *)
  FUEL_CELLFT-02_ALARM_HI := 0.0 ;  (* expected-zero state: any positive PV alarms )

  (* FLOW control loop - set-point from the graph basis *)
  FUEL_CELLFT-03_SP := 0.01 ;  (* graph basis: IA-FC-LEACH normal 0.01 L/h )
  FB_PI_FUEL_CELLFT-03( PV := FUEL_CELLFT-03_PV, SP := FUEL_CELLFT-03_SP );  (* PI per AQS-CTL-002; GAIN/KI entered at commissioning from the step test (AQS-COM-001 sec. 3), anti-windup clamp per this FB *)
  FUEL_CELLFT-03_ALARM_HI := 0.011000000000000001 ;  (* SP x 1.1 margin, A-M-188 margin class *)
  FUEL_CELLFT-03_ALARM_LO := 0.009000000000000001 ;

  (* PRESSURE monitoring block - indication, no set-point invented )
  FB_AI_FUEL_CELLPT-01( PV := FUEL_CELLPT-01_PV );
  FUEL_CELLPT-01_ALARM_HI := 9.0 ;  (* 90 % of span, registered LSH convention )

  (* TEMPERATURE monitoring block - indication, no set-point invented )
  FB_AI_FUEL_CELLTE-01( PV := FUEL_CELLTE-01_PV );
  FUEL_CELLTE-01_ALARM_HI := 135.0 ;  (* 90 % of span, registered LSH convention )

  (* PRESSURE monitoring block - indication, no set-point invented )
  FB_AI_PV_ARRAYPT-01( PV := PV_ARRAYPT-01_PV );
  PV_ARRAYPT-01_ALARM_HI := 9.0 ;  (* 90 % of span, registered LSH convention )

  (* TEMPERATURE monitoring block - indication, no set-point invented )
  FB_AI_PV_ARRAYTE-01( PV := PV_ARRAYTE-01_PV );
  PV_ARRAYTE-01_ALARM_HI := 135.0 ;  (* 90 % of span, registered LSH convention )

  (* PRESSURE monitoring block - indication, no set-point invented )
  FB_AI_RECTIFIERPT-01( PV := RECTIFIERPT-01_PV );
  RECTIFIERPT-01_ALARM_HI := 9.0 ;  (* 90 % of span, registered LSH convention )

  (* TEMPERATURE monitoring block - indication, no set-point invented )
  FB_AI_RECTIFIERTE-01( PV := RECTIFIERTE-01_PV );
  RECTIFIERTE-01_ALARM_HI := 135.0 ;  (* 90 % of span, registered LSH convention )

  (* FLOW control loop - set-point from the graph basis *)
  ZNBR2_BR2_REGENFT-01_SP := 33.48 ;  (* graph basis: S69B normal 33.48 L/h )
  FB_PI_ZNBR2_BR2_REGENFT-01( PV := ZNBR2_BR2_REGENFT-01_PV, SP := ZNBR2_BR2_REGENFT-01_SP );  (* PI per AQS-CTL-002; GAIN/KI entered at commissioning from the step test (AQS-COM-001 sec. 3), anti-windup clamp per this FB *)
  ZNBR2_BR2_REGENFT-01_ALARM_HI := 36.828 ;  (* SP x 1.1 margin, A-M-188 margin class *)
  ZNBR2_BR2_REGENFT-01_ALARM_LO := 30.131999999999998 ;

  (* LEVEL monitoring block - indication, no set-point invented )
  FB_AI_ZNBR2_BR2_REGENLT-01( PV := ZNBR2_BR2_REGENLT-01_PV );
  ZNBR2_BR2_REGENLT-01_ALARM_HI := 90.0 ;  (* 90 % of span, registered LSH convention )

  (* PRESSURE monitoring block - indication, no set-point invented )
  FB_AI_ZNBR2_BR2_REGENPT-01( PV := ZNBR2_BR2_REGENPT-01_PV );
  ZNBR2_BR2_REGENPT-01_ALARM_HI := 9.0 ;  (* 90 % of span, registered LSH convention )

  (* TEMPERATURE monitoring block - indication, no set-point invented )
  FB_AI_ZNBR2_BR2_REGENTE-01( PV := ZNBR2_BR2_REGENTE-01_PV );
  ZNBR2_BR2_REGENTE-01_ALARM_HI := 135.0 ;  (* 90 % of span, registered LSH convention )

  (* TEMPERATURE monitoring block - indication, no set-point invented )
  FB_AI_EXT_HALLTE-01( PV := EXT_HALLTE-01_PV );
  EXT_HALLTE-01_ALARM_HI := 135.0 ;  (* 90 % of span, registered LSH convention )

  (* PRESSURE monitoring block - indication, no set-point invented )
  FB_AI_LIO_BATPT-01( PV := LIO_BATPT-01_PV );
  LIO_BATPT-01_ALARM_HI := 630.0 ;  (* 90 % of span, registered LSH convention )

END_PROGRAM
